(* IEC 61131-3 sources: plcassist-cli/packages/volt-lsp-iec/test-corpus/bakon-nano/Device/Plc Logic/Application/Library Manager/L_UBUP_BasicUtilities, 147 files *)

(* ---- L_UBUP_INTERNAL.gvl ---- *)
VAR_GLOBAL
	ONLINECHANGEDETECTION : L_UBUP_OnlineChangeDetection;
	LMJOBADMINSTRATION : L_UBUP_JobAdminstration;
	G_FBPOOLQUEUE : L_UBUP_JobPoolQueue;
	G_ILOWESTREQUESTPRIO : INT := DWORD_TO_INT(16#7FFF);
	G_DWCALLIDUNASSIGNED : DWORD := 4711;
	CDIENUMSTARTVALUE : DINT := 10000;
END_VAR

(* ---- L_UBUP_IACTIONPROVIDER.itf ---- *)
INTERFACE L_UBUP_IACTIONPROVIDER
END_INTERFACE

METHOD CYCLICACTION
VAR_INPUT
	ITFTIMINGCONTROLLER : L_UBUP_ITimingController;
END_VAR
VAR_OUTPUT
	XCOMPLETE : BOOL;
	XABORT : BOOL;
	IERRORID : INT;
END_VAR
END_METHOD

METHOD FINALIZEACTION
VAR_INPUT
	XABORTPROPOSED : BOOL;
	IERRORIDPROPOSED : INT;
END_VAR
VAR_OUTPUT
	XCOMPLETE : BOOL;
	XABORT : BOOL;
	IERRORID : INT;
END_VAR
END_METHOD

METHOD RESETACTION
VAR_OUTPUT
	XCOMPLETE : BOOL;
END_VAR
END_METHOD

METHOD STARTACTION
VAR_OUTPUT
	XCOMPLETE : BOOL;
	IERRORID : INT;
END_VAR
END_METHOD

(* ---- L_UBUP_IAFTERREADINPUTS.itf ---- *)
INTERFACE L_UBUP_IAFTERREADINPUTS
END_INTERFACE

METHOD AFTERREADINPUTS : INT
END_METHOD

(* ---- L_UBUP_IAFTERREADINPUTSEXIT.itf ---- *)
INTERFACE L_UBUP_IAFTERREADINPUTSEXIT
END_INTERFACE

METHOD AFTERREADINPUTSEXIT : INT
END_METHOD

(* ---- L_UBUP_IAFTERWRITEOUTPUTS.itf ---- *)
INTERFACE L_UBUP_IAFTERWRITEOUTPUTS
END_INTERFACE

METHOD AFTERWRITEOUTPUTS : INT
END_METHOD

(* ---- L_UBUP_IAFTERWRITEOUTPUTSEXIT.itf ---- *)
INTERFACE L_UBUP_IAFTERWRITEOUTPUTSEXIT
END_INTERFACE

METHOD AFTERWRITEOUTPUTSEXIT : INT
END_METHOD

(* ---- L_UBUP_IALLOCPOINTADRPROVIDER.itf ---- *)
INTERFACE L_UBUP_IALLOCPOINTADRPROVIDER
END_INTERFACE

METHOD ALLOCPOINTADR
VAR_OUTPUT
	IERRORID : INT;
END_VAR
END_METHOD

(* ---- L_UBUP_IALTERNATIVEREQUESTBYFAILEDCONDITION.itf ---- *)
INTERFACE L_UBUP_IALTERNATIVEREQUESTBYFAILEDCONDITION
END_INTERFACE

METHOD HANDLEREJECTEDREQUEST : BOOL
VAR_INPUT
	ITFREQUESTANNOUNCED : L_UBUP_IRequest;
END_VAR
VAR_OUTPUT
	ITFALTERNATIVEREQUEST : L_UBUP_IRequest;
END_VAR
END_METHOD

(* ---- L_UBUP_IBEFOREREADINPUTS.itf ---- *)
INTERFACE L_UBUP_IBEFOREREADINPUTS
END_INTERFACE

METHOD BEFOREREADINPUTS : INT
END_METHOD

(* ---- L_UBUP_IBEFOREREADINPUTSENTRY.itf ---- *)
INTERFACE L_UBUP_IBEFOREREADINPUTSENTRY
END_INTERFACE

METHOD BEFOREREADINPUTSENTRY : INT
END_METHOD

(* ---- L_UBUP_IBEFOREWRITEOUTPUTS.itf ---- *)
INTERFACE L_UBUP_IBEFOREWRITEOUTPUTS
END_INTERFACE

METHOD BEFOREWRITEOUTPUTS : INT
END_METHOD

(* ---- L_UBUP_IBEFOREWRITEOUTPUTSENTRY.itf ---- *)
INTERFACE L_UBUP_IBEFOREWRITEOUTPUTSENTRY
END_INTERFACE

METHOD BEFOREWRITEOUTPUTSENTRY : INT
END_METHOD

(* ---- L_UBUP_IBREAKPOINT.itf ---- *)
INTERFACE L_UBUP_IBREAKPOINT
END_INTERFACE

METHOD BREAKPOINT : INT
END_METHOD

(* ---- L_UBUP_ICATEGORY.itf ---- *)
INTERFACE L_UBUP_ICATEGORY
END_INTERFACE

METHOD CLASSIFY : BOOL
VAR_INPUT
	ECATEGORY : DINT;
END_VAR
END_METHOD

(* ---- L_UBUP_ICHECKER.itf ---- *)
INTERFACE L_UBUP_ICHECKER
END_INTERFACE

METHOD PERFORMCHECK : BOOL
VAR_INPUT
	WCONTEXT : DWORD;
END_VAR
END_METHOD

(* ---- L_UBUP_ICOMMAND.itf ---- *)
INTERFACE L_UBUP_ICOMMAND
END_INTERFACE

METHOD UPDATECOMMANDDATA : BOOL
VAR_INPUT
	DWCALLID : DWORD;
	XCONTINUOUSUPDATE : BOOL;
END_VAR
VAR_IN_OUT
	SCCOMMAND : L_UBUP_CommandData;
END_VAR
END_METHOD

(* ---- L_UBUP_ICOMPARER.itf ---- *)
INTERFACE L_UBUP_ICOMPARER
END_INTERFACE

METHOD COMPARE : DINT
VAR_INPUT
	DWARRIDX1 : DWORD;
	DWARRIDX2 : DWORD;
END_VAR
END_METHOD

(* ---- L_UBUP_ICONDITION.itf ---- *)
INTERFACE L_UBUP_ICONDITION
END_INTERFACE

METHOD VERIFY : BOOL
VAR_OUTPUT
	XCONDITIONERROR : BOOL;
	EERRORIDPROPOSED : L_IE1P_Error;
END_VAR
END_METHOD

(* ---- L_UBUP_ICRITICALSECTION.itf ---- *)
INTERFACE L_UBUP_ICRITICALSECTION
END_INTERFACE

METHOD LOCK : BOOL
END_METHOD

METHOD LOCKSTATE : BOOL
END_METHOD

METHOD UNLOCK : BOOL
END_METHOD

(* ---- L_UBUP_IEXCEPTION.itf ---- *)
INTERFACE L_UBUP_IEXCEPTION
END_INTERFACE

METHOD EXCEPTION : INT
END_METHOD

(* ---- L_UBUP_IFBPOOL.itf ---- *)
INTERFACE L_UBUP_IFBPOOL
END_INTERFACE

METHOD FREEINSTANCE : BOOL
VAR_INPUT
	ITFINSTANCE : L_UBUP_IPoolInstance;
	XWHANDLE : __XWORD;
END_VAR
END_METHOD

METHOD GETCAPACITY : BOOL
VAR_INPUT
	ECLASSID : DINT;
END_VAR
VAR_OUTPUT
	DWCAPACITY : DWORD;
END_VAR
END_METHOD

METHOD QUERYINSTANCE : BOOL
VAR_INPUT
	ECLASSID : DINT;
END_VAR
VAR_IN_OUT
	ITFINSTANCE : L_UBUP_IPoolInstance;
END_VAR
END_METHOD

(* ---- L_UBUP_IINSTANCE.itf ---- *)
INTERFACE L_UBUP_IINSTANCE
END_INTERFACE

(* ---- L_UBUP_IINSTANCELIST.itf ---- *)
INTERFACE L_UBUP_IINSTANCELIST
END_INTERFACE

METHOD APPENDPROXY : BOOL
VAR_INPUT
	ITFINSTANCELISTITEM : L_UBUP_IInstanceListProxy;
END_VAR
END_METHOD

(* ---- L_UBUP_IINSTANCELISTPASSENGER.itf ---- *)
INTERFACE L_UBUP_IINSTANCELISTPASSENGER
END_INTERFACE

(* ---- L_UBUP_IINSTANCELISTPROXY.itf ---- *)
INTERFACE L_UBUP_IINSTANCELISTPROXY
END_INTERFACE

(* ---- L_UBUP_IITERATOR.itf ---- *)
INTERFACE L_UBUP_IITERATOR
END_INTERFACE

METHOD NEXT : DWORD
END_METHOD

METHOD PREV : DWORD
END_METHOD

METHOD REWIND
VAR_OUTPUT
	DWARRAYIDXSTART : DWORD;
END_VAR
END_METHOD

(* ---- L_UBUP_IJOB.itf ---- *)
INTERFACE L_UBUP_IJOB
END_INTERFACE

METHOD EXPAND : BOOL
VAR_INPUT
	ITFSENDER : L_UBUP_ICommand;
	DWCALLID : DWORD;
END_VAR
VAR_OUTPUT
	EERRORID : L_IE1P_Error;
END_VAR
END_METHOD

METHOD HANDOVERRESOURCE : BOOL
VAR_INPUT
	ITFRESOURCE : L_UBUP_IUnknown;
END_VAR
END_METHOD

METHOD LINK : BOOL
VAR_INPUT
	ITFJOB : L_UBUP_IJob;
	XPREV : BOOL;
END_VAR
VAR_OUTPUT
	EERRORID : L_IE1P_Error;
END_VAR
END_METHOD

METHOD RELEASE
END_METHOD

(* ---- L_UBUP_IJOBACTION.itf ---- *)
INTERFACE L_UBUP_IJOBACTION
END_INTERFACE

METHOD ABORT
END_METHOD

METHOD CYCLE
VAR_OUTPUT
	ESTATE : L_UBUP_JobState;
	EERRORID : L_IE1P_Error;
END_VAR
END_METHOD

METHOD FINISH
END_METHOD

METHOD UPDATEREPORTDATA : BOOL
VAR_INPUT
	DWCALLID : DWORD;
END_VAR
VAR_IN_OUT
	SCREPORT : L_UBUP_ReportData;
END_VAR
END_METHOD

METHOD UPDATEREPORTRECEIVER : BOOL
VAR_INPUT
	ITFJOBREPORT : L_UBUP_IJobReport;
END_VAR
END_METHOD

(* ---- L_UBUP_IJOBCOLLECTION.itf ---- *)
INTERFACE L_UBUP_IJOBCOLLECTION
END_INTERFACE

METHOD GETJOB : BOOL
VAR_INPUT
	DWARRIDX : DWORD;
END_VAR
VAR_OUTPUT
	ITFJOB : L_UBUP_IJob;
END_VAR
END_METHOD

(* ---- L_UBUP_IJOBRECEIVER.itf ---- *)
INTERFACE L_UBUP_IJOBRECEIVER
END_INTERFACE

METHOD INSERT : BOOL
VAR_INPUT
	ITFJOB : L_UBUP_IJob;
END_VAR
END_METHOD

METHOD UNPLUGLISTENER : BOOL
VAR_INPUT
	ITFLISTENER : L_UBUP_IJobReceiverListener;
END_VAR
END_METHOD

METHOD ANNOUNCELISTENER : BOOL
VAR_INPUT
	ITFLISTENER : L_UBUP_IJobReceiverListener;
END_VAR
END_METHOD

(* ---- L_UBUP_IJOBRECEIVERLISTENER.itf ---- *)
INTERFACE L_UBUP_IJOBRECEIVERLISTENER
END_INTERFACE

METHOD LISTENAFTERCYCLE
VAR_INPUT
	ITFJOB : L_UBUP_IJob;
END_VAR
END_METHOD

METHOD LISTENINSERT
VAR_INPUT
	ITFJOB : L_UBUP_IJob;
	XSUCCEEDED : BOOL;
END_VAR
END_METHOD

(* ---- L_UBUP_IJOBREPORT.itf ---- *)
INTERFACE L_UBUP_IJOBREPORT
END_INTERFACE

METHOD RECEIVEREPORT
VAR_INPUT
	ITFJOB : L_UBUP_IJob;
END_VAR
END_METHOD

(* ---- L_UBUP_ILIST.itf ---- *)
INTERFACE L_UBUP_ILIST
END_INTERFACE

(* ---- L_UBUP_ILISTCONTROL.itf ---- *)
INTERFACE L_UBUP_ILISTCONTROL
END_INTERFACE

METHOD APPEND : BOOL
VAR_OUTPUT
	DWARRIDX : DWORD;
END_VAR
END_METHOD

METHOD GETARRIDXOF : DWORD
VAR_INPUT
	DWPOSITION : DWORD;
END_VAR
END_METHOD

METHOD GETMAX : DWORD
VAR_INPUT
	ITFCOMPARER : L_UBUP_IComparer;
END_VAR
END_METHOD

METHOD GETPOSITIONOF : DWORD
VAR_INPUT
	DWARRIDX : DWORD;
END_VAR
END_METHOD

METHOD INSERTAFTER : BOOL
VAR_INPUT
	DWARRIDX : DWORD;
END_VAR
VAR_OUTPUT
	DWNEXTIDX : DWORD;
END_VAR
END_METHOD

METHOD INSERTBEFORE : BOOL
VAR_INPUT
	DWARRIDX : DWORD;
END_VAR
VAR_OUTPUT
	DWPREVIDX : DWORD;
END_VAR
END_METHOD

METHOD REMOVE : BOOL
VAR_INPUT
	DWARRIDX : DWORD;
END_VAR
END_METHOD

METHOD SHIFTNEXT : BOOL
VAR_INPUT
	DWARRIDX : DWORD;
END_VAR
END_METHOD

METHOD SHIFTPREV : BOOL
VAR_INPUT
	DWARRIDX : DWORD;
END_VAR
END_METHOD

METHOD SORT : BOOL
VAR_INPUT
	ITFCOMPARER : L_UBUP_IComparer;
END_VAR
END_METHOD

METHOD SWAP : BOOL
VAR_INPUT
	DWARRIDX1 : DWORD;
	DWARRIDX2 : DWORD;
END_VAR
END_METHOD

METHOD TRYAPPEND : BOOL
VAR_INPUT
	DWARRIDX : DWORD;
END_VAR
END_METHOD

(* ---- L_UBUP_ILMDATA.itf ---- *)
INTERFACE L_UBUP_ILMDATA
END_INTERFACE

METHOD ABORT : UDINT
END_METHOD

METHOD EXECUTE : UDINT
END_METHOD

(* ---- L_UBUP_ILOCKABLE.itf ---- *)
INTERFACE L_UBUP_ILOCKABLE
END_INTERFACE

METHOD LOCK : BOOL
END_METHOD

METHOD LOCKSTATE : BOOL
END_METHOD

METHOD UNLOCK : BOOL
END_METHOD

(* ---- L_UBUP_IMAPOUTPUTSPROVIDER.itf ---- *)
INTERFACE L_UBUP_IMAPOUTPUTSPROVIDER
END_INTERFACE

METHOD MAPOUTPUTS
END_METHOD

(* ---- L_UBUP_IMAPSTATE.itf ---- *)
INTERFACE L_UBUP_IMAPSTATE
END_INTERFACE

(* ---- L_UBUP_IMEMORYCONSUMER.itf ---- *)
INTERFACE L_UBUP_IMEMORYCONSUMER
END_INTERFACE

METHOD EVALMEMORYPROVIDER
VAR_INPUT
	ITFMEMORYPROVIDER : L_UBUP_IMemoryProvider;
END_VAR
END_METHOD

(* ---- L_UBUP_IMEMORYPROVIDER.itf ---- *)
INTERFACE L_UBUP_IMEMORYPROVIDER
END_INTERFACE

METHOD REGISTERCONSUMER
VAR_INPUT
	ITFMEMORYCONSUMER : L_UBUP_IMemoryConsumer;
END_VAR
END_METHOD

(* ---- L_UBUP_IMONITORSTATESERVER.itf ---- *)
INTERFACE L_UBUP_IMONITORSTATESERVER
END_INTERFACE

METHOD MONITORCASE
VAR_INPUT
	ECASE : L_UBUP_StateHandleCase;
END_VAR
END_METHOD

METHOD MONITORREQUEST : INT
VAR_INPUT
	ITFREQUEST : L_UBUP_IRequest;
END_VAR
END_METHOD

METHOD MONITORREQUESTANNOUNCED : INT
VAR_INPUT
	ITFREQUESTANNOUNCED : L_UBUP_IRequest;
	ITFREQUESTALTERNATIVE : L_UBUP_IRequest := 0;
	ITFREQUESTACTIVE : L_UBUP_IRequest;
END_VAR
END_METHOD

(* ---- L_UBUP_IOBJECT.itf ---- *)
INTERFACE L_UBUP_IOBJECT
END_INTERFACE

METHOD CALL_INIT : BOOL
END_METHOD

METHOD SETNEXT : BOOL
VAR_INPUT
	ITFOBJECT : L_UBUP_IObject;
END_VAR
END_METHOD

METHOD SETPREV : BOOL
VAR_INPUT
	ITFOBJECT : L_UBUP_IObject;
END_VAR
END_METHOD

(* ---- L_UBUP_IOBJECTQUEUE.itf ---- *)
INTERFACE L_UBUP_IOBJECTQUEUE
END_INTERFACE

METHOD DEQUEUE : BOOL
END_METHOD

METHOD ENQUEUE : BOOL
VAR_INPUT
	ITFOBJECT : L_UBUP_IObject;
END_VAR
END_METHOD

METHOD REMOVE : BOOL
VAR_INPUT
	ITFOBJECT : L_UBUP_IObject;
END_VAR
END_METHOD

(* ---- L_UBUP_IPLCOPENSTATUS.itf ---- *)
INTERFACE L_UBUP_IPLCOPENSTATUS
END_INTERFACE

METHOD GET_EERRORID : L_IE1P_Error
END_METHOD

METHOD GET_XACTIVE : BOOL
END_METHOD

METHOD GET_XBUSY : BOOL
END_METHOD

METHOD GET_XCOMMANDABORTED : BOOL
END_METHOD

METHOD GET_XDONE : BOOL
END_METHOD

METHOD GET_XINITIAL : BOOL
END_METHOD

(* ---- L_UBUP_IPOINTERCOLLECTION.itf ---- *)
INTERFACE L_UBUP_IPOINTERCOLLECTION
END_INTERFACE

METHOD GETPOINTER : BOOL
VAR_INPUT
	DWARRIDX : DWORD;
END_VAR
VAR_OUTPUT
	PBYTE : POINTER TO BYTE;
END_VAR
END_METHOD

(* ---- L_UBUP_IPOOLINSTANCE.itf ---- *)
INTERFACE L_UBUP_IPOOLINSTANCE
END_INTERFACE

METHOD FREE : BOOL
END_METHOD

METHOD OCCUPY : BOOL
VAR_INPUT
	ITFOWNER : L_UBUP_IFBPool;
	XWHANDLE : __XWORD;
END_VAR
END_METHOD

(* ---- L_UBUP_IQUEUE.itf ---- *)
INTERFACE L_UBUP_IQUEUE
END_INTERFACE

METHOD DEQUEUE : BOOL
END_METHOD

METHOD ENQUEUE : BOOL
END_METHOD

METHOD GETEMPTY : BOOL
VAR_OUTPUT
	PBYTE : POINTER TO BYTE;
	DWSIZE : DWORD;
END_VAR
END_METHOD

METHOD GETPEEK : BOOL
VAR_OUTPUT
	PBYTE : POINTER TO BYTE;
	DWSIZE : DWORD;
END_VAR
END_METHOD

METHOD RESET : BOOL
END_METHOD

(* ---- L_UBUP_IREADINPUTSEXIT.itf ---- *)
INTERFACE L_UBUP_IREADINPUTSEXIT
END_INTERFACE

METHOD READINPUTSEXIT : INT
END_METHOD

(* ---- L_UBUP_IREFCOUNTER.itf ---- *)
INTERFACE L_UBUP_IREFCOUNTER
END_INTERFACE

METHOD DECCOUNTER : DINT
END_METHOD

METHOD INCCOUNTER : DINT
END_METHOD

(* ---- L_UBUP_IREQUEST.itf ---- *)
INTERFACE L_UBUP_IREQUEST
END_INTERFACE

METHOD CONFIRM : INT
VAR_IN_OUT
	IREQUEST : L_UBUP_IRequest;
END_VAR
END_METHOD

METHOD FORCESTATEENTRY : BOOL
END_METHOD

(* ---- L_UBUP_ISTATECLIENT.itf ---- *)
INTERFACE L_UBUP_ISTATECLIENT
END_INTERFACE

METHOD CALLFBS
VAR_INPUT
	ECASE : L_UBUP_StateHandleCase;
END_VAR
END_METHOD

METHOD CALLSTATE
VAR_INPUT
	ITFSTATESERVER : L_UBUP_IStateServer;
	ISTATE : INT;
	ECASE : L_UBUP_StateHandleCase;
END_VAR
END_METHOD

METHOD CHECKTRANSITION
VAR_INPUT
	ITFSTATESERVER : L_UBUP_IStateServer;
END_VAR
END_METHOD

METHOD DISABLECLIENT : BOOL
VAR_INPUT
	XFIRSTCALL : BOOL;
END_VAR
END_METHOD

METHOD ENABLECLIENT : BOOL
VAR_INPUT
	XFIRSTCALL : BOOL;
END_VAR
END_METHOD

METHOD FINALIZECYCLE
END_METHOD

METHOD LEAVESTATE
END_METHOD

METHOD PREPARECYCLE
END_METHOD

METHOD PREPARESTATECHANGE
END_METHOD

METHOD STIMULATETRANSITION
VAR_INPUT
	ECASE : L_UBUP_StateHandleCase;
END_VAR
END_METHOD

METHOD UPDATECONDITIONERROR : BOOL
VAR_INPUT
	ITFREQUEST : L_UBUP_IRequest;
END_VAR
END_METHOD

(* ---- L_UBUP_ISTATECLIENTDECORATOR.itf ---- *)
INTERFACE L_UBUP_ISTATECLIENTDECORATOR
END_INTERFACE

METHOD EXTENDEDCALLFBS
VAR_INPUT
	ECASE : L_UBUP_StateHandleCase;
END_VAR
END_METHOD

METHOD EXTENDEDCALLSTATE
VAR_INPUT
	ITFBASE : L_UBUP_IStateClient;
	ITFSTATESERVER : L_UBUP_IStateServer;
	ISTATE : INT;
	ECASE : L_UBUP_StateHandleCase;
END_VAR
END_METHOD

METHOD EXTENDEDCHECKTRANSITION
VAR_INPUT
	ITFSTATESERVER : L_UBUP_IStateServer;
END_VAR
END_METHOD

METHOD EXTENDEDDISABLECLIENT : BOOL
VAR_INPUT
	XFIRSTCALL : BOOL;
END_VAR
END_METHOD

METHOD EXTENDEDENABLECLIENT : BOOL
VAR_INPUT
	XFIRSTCALL : BOOL;
END_VAR
END_METHOD

METHOD EXTENDEDFINALIZECYCLE
END_METHOD

METHOD EXTENDEDPREPARECYCLE
END_METHOD

METHOD EXTENDEDPREPARESTATECHANGE
END_METHOD

METHOD EXTENDEDSTIMULATETRANSITION
VAR_INPUT
	ECASE : L_UBUP_StateHandleCase;
END_VAR
END_METHOD

(* ---- L_UBUP_ISTATESERVER.itf ---- *)
INTERFACE L_UBUP_ISTATESERVER
END_INTERFACE

METHOD ANNOUNCENEWREQUEST
END_METHOD

METHOD FREEZEREQUEST
VAR_INPUT
	EERRORIDBYBLOCKEFREEZEREQUEST : L_IE1P_Error;
END_VAR
END_METHOD

METHOD ISACTIVE : BOOL
VAR_INPUT
	ITFREQUEST : L_UBUP_IRequest;
END_VAR
END_METHOD

METHOD REQUESTS : INT
VAR_INPUT
	ITFREQUEST : L_UBUP_IRequest;
END_VAR
END_METHOD

METHOD UNFREEZEREQUEST : BOOL
END_METHOD

METHOD VERIFYFREEZEREQUEST : BOOL
VAR_INPUT
	ITFREQUEST : L_UBUP_IRequest;
END_VAR
VAR_OUTPUT
	XCONDITIONERROR : BOOL;
	EERRORIDPROPOSED : L_IE1P_Error;
END_VAR
END_METHOD

(* ---- L_UBUP_ISTRINGCOLLECTION.itf ---- *)
INTERFACE L_UBUP_ISTRINGCOLLECTION
END_INTERFACE

METHOD GETSTRING : BOOL
VAR_INPUT
	DWARRIDX : DWORD;
END_VAR
VAR_OUTPUT
	STVALUE : STRING(255);
END_VAR
END_METHOD

(* ---- L_UBUP_ITIMINGCONTROLLER.itf ---- *)
INTERFACE L_UBUP_ITIMINGCONTROLLER
END_INTERFACE

METHOD CHECKTIMING
VAR_OUTPUT
	XTIMEOUT : BOOL;
	XTIMELIMIT : BOOL;
END_VAR
END_METHOD

METHOD STARTINVOCATIONTIMER
END_METHOD

METHOD STARTOPERATIONTIMER
END_METHOD

(* ---- L_UBUP_IUNKNOWN.itf ---- *)
INTERFACE L_UBUP_IUNKNOWN
END_INTERFACE

METHOD REQUESTINTERFACE : BOOL
VAR_INPUT
	ID : DINT;
	PITFUNKNOWN : POINTER TO L_UBUP_IUnknown;
END_VAR
END_METHOD

(* ---- L_UBUP_IWRITEOUTPUTSENTRY.itf ---- *)
INTERFACE L_UBUP_IWRITEOUTPUTSENTRY
END_INTERFACE

METHOD WRITEOUTPUTSENTRY : INT
END_METHOD

(* ---- GETBOOLEANPROPERTY.fun ---- *)
FUNCTION GETBOOLEANPROPERTY : BOOL
VAR_INPUT
	STKEY : WSTRING;
END_VAR
END_FUNCTION

(* ---- GETCOMPANY.fun ---- *)
FUNCTION GETCOMPANY : WSTRING
END_FUNCTION

(* ---- GETNUMBERPROPERTY.fun ---- *)
FUNCTION GETNUMBERPROPERTY : DINT
VAR_INPUT
	STKEY : WSTRING;
END_VAR
END_FUNCTION

(* ---- GETTEXTPROPERTY.fun ---- *)
FUNCTION GETTEXTPROPERTY : WSTRING
VAR_INPUT
	STKEY : WSTRING;
END_VAR
END_FUNCTION

(* ---- GETTEXTPROPERTY2.fun ---- *)
FUNCTION GETTEXTPROPERTY2 : POINTER TO WSTRING
VAR_INPUT
	STKEY : WSTRING;
END_VAR
END_FUNCTION

(* ---- GETTITLE.fun ---- *)
FUNCTION GETTITLE : WSTRING
END_FUNCTION

(* ---- GETVERSION.fun ---- *)
FUNCTION GETVERSION : VERSION
END_FUNCTION

(* ---- GETVERSIONPROPERTY.fun ---- *)
FUNCTION GETVERSIONPROPERTY : VERSION
VAR_INPUT
	STKEY : WSTRING;
END_VAR
END_FUNCTION

(* ---- L_UBUP_CREATECALLID.fun ---- *)
FUNCTION L_UBUP_CREATECALLID : DWORD
END_FUNCTION

(* ---- L_UBUP_CREATEOBJECTID.fun ---- *)
FUNCTION L_UBUP_CREATEOBJECTID : DWORD
END_FUNCTION

(* ---- L_UBUP_FILEADDRESS.fun ---- *)
FUNCTION L_UBUP_FILEADDRESS : STRING(255)
END_FUNCTION

(* ---- L_UBUP_GETTASKCYCLE.fun ---- *)
FUNCTION L_UBUP_GETTASKCYCLE : LREAL
VAR_INPUT
	LRCYCLETIMEIN : LREAL;
END_VAR
END_FUNCTION

(* ---- L_UBUP_GETTASKINFO.fun ---- *)
FUNCTION L_UBUP_GETTASKINFO : BOOL
VAR_OUTPUT
	ITASKINDEX : INT;
	HTASK : RTS_IEC_HANDLE;
	HIECTASK : RTS_IEC_HANDLE;
	PSCSYSTASKINFO : POINTER TO SYS_TASK_INFO;
	UDIOSPRIORITY : UDINT;
	UDIPRIORITY : UDINT;
	UDITASKINTERVAL : UDINT;
END_VAR
END_FUNCTION

(* ---- L_UBUP_ISLENZETARGET.fun ---- *)
FUNCTION L_UBUP_ISLENZETARGET : BOOL
VAR_OUTPUT
	DWVENDORID : DWORD;
END_VAR
END_FUNCTION

(* ---- L_UBUP_ISONLINECHANGEACTIVE.fun ---- *)
FUNCTION L_UBUP_ISONLINECHANGEACTIVE : BOOL
END_FUNCTION

(* ---- L_UBUP_LMDATAMANAGERINSERTDATA.fun ---- *)
FUNCTION L_UBUP_LMDATAMANAGERINSERTDATA : BOOL
VAR_INPUT
	ITFLMDATA : L_UBUP_ILMData;
END_VAR
END_FUNCTION

(* ---- L_UBUP_LOCALDATEANDTIME.fun ---- *)
FUNCTION L_UBUP_LOCALDATEANDTIME : BOOL
VAR_OUTPUT
	UIYEAR : UINT;
	UIMONTH : UINT;
	UIDAY : UINT;
	UIHOUR : UINT;
	UIMINUTE : UINT;
	UISECOND : UINT;
	UIMILLISECONDS : UINT;
	UIWEEKDAY : UINT;
	DATDATE : DATE;
	TODTIME : TIME_OF_DAY;
END_VAR
END_FUNCTION

(* ---- L_UBUP_QUERY_IJOB_ALL.fun ---- *)
FUNCTION L_UBUP_QUERY_IJOB_ALL : BOOL
VAR_INPUT
	ITFJOB : L_UBUP_IJob;
END_VAR
VAR_OUTPUT
	ITFINSTANCE : L_UBUP_IPoolInstance;
	ITFSTATECLIENT : L_UBUP_IStateClient;
	ITFPLCOPENSTATUS : L_UBUP_IPLCOpenStatus;
END_VAR
END_FUNCTION

(* ---- L_UBUP_QUERY_IJOB_IINSTANCE.fun ---- *)
FUNCTION L_UBUP_QUERY_IJOB_IINSTANCE : BOOL
VAR_INPUT
	ITFJOB : L_UBUP_IJob;
END_VAR
VAR_OUTPUT
	ITFINSTANCE : L_UBUP_IPoolInstance;
END_VAR
END_FUNCTION

(* ---- L_UBUP_QUERY_IJOB_IPLCOPENSTATUS.fun ---- *)
FUNCTION L_UBUP_QUERY_IJOB_IPLCOPENSTATUS : BOOL
VAR_INPUT
	ITFJOB : L_UBUP_IJob;
END_VAR
VAR_OUTPUT
	ITFPLCOPENSTATUS : L_UBUP_IPLCOpenStatus;
END_VAR
END_FUNCTION

(* ---- L_UBUP_SYMBOLCONFIGREADNUMVAR.fun ---- *)
FUNCTION L_UBUP_SYMBOLCONFIGREADNUMVAR : BOOL
VAR_INPUT
	SVARIABLENAME : STRING;
END_VAR
VAR_OUTPUT
	SCVARIABLE : L_UBUP_Variable;
END_VAR
END_FUNCTION

(* ---- L_UBUP_SYMBOLCONFIGREADSTRINGVAR.fun ---- *)
FUNCTION L_UBUP_SYMBOLCONFIGREADSTRINGVAR : BOOL
VAR_INPUT
	SVARIABLENAME : STRING;
END_VAR
VAR_OUTPUT
	SVALUE : STRING;
END_VAR
END_FUNCTION

(* ---- L_UBUP_SYMBOLCONFIGREADVAR.fun ---- *)
FUNCTION L_UBUP_SYMBOLCONFIGREADVAR : BOOL
VAR_INPUT
	SVARIABLENAME : STRING;
END_VAR
VAR_OUTPUT
	SCVARIABLE : L_UBUP_Variable;
END_VAR
END_FUNCTION

(* ---- L_UBUP_SYMBOLCONFIGREADVARASDWORD.fun ---- *)
FUNCTION L_UBUP_SYMBOLCONFIGREADVARASDWORD : BOOL
VAR_INPUT
	SVARIABLENAME : STRING;
END_VAR
VAR_OUTPUT
	DWVALUE : DWORD;
END_VAR
END_FUNCTION

(* ---- L_UBUP_SYMBOLCONFIGREADVARASLINT.fun ---- *)
FUNCTION L_UBUP_SYMBOLCONFIGREADVARASLINT : BOOL
VAR_INPUT
	SVARIABLENAME : STRING;
END_VAR
VAR_OUTPUT
	LIVALUE : LINT;
END_VAR
END_FUNCTION

(* ---- L_UBUP_SYMBOLCONFIGREADVARASLREAL.fun ---- *)
FUNCTION L_UBUP_SYMBOLCONFIGREADVARASLREAL : BOOL
VAR_INPUT
	SVARIABLENAME : STRING;
END_VAR
VAR_OUTPUT
	LRVALUE : LREAL;
END_VAR
END_FUNCTION

(* ---- L_UBUP_SYMBOLCONFIGREADVARASWORD.fun ---- *)
FUNCTION L_UBUP_SYMBOLCONFIGREADVARASWORD : BOOL
VAR_INPUT
	SVARIABLENAME : STRING;
END_VAR
VAR_OUTPUT
	WVALUE : WORD;
END_VAR
END_FUNCTION

(* ---- L_UBUP_SYMBOLCONFIGSYMBOLEXISTS.fun ---- *)
FUNCTION L_UBUP_SYMBOLCONFIGSYMBOLEXISTS : BOOL
VAR_INPUT
	SVARIABLENAME : STRING;
END_VAR
END_FUNCTION

(* ---- GLOBALTEXTLIST.fb ---- *)
FUNCTION_BLOCK GLOBALTEXTLIST
VAR
	M_TEXTLISTFILE : STRING(255);
	_STNAMESPACE : STRING;
END_VAR
END_FUNCTION_BLOCK

(* ---- L_UBUP_BEHAVIOURMODEL.fb ---- *)
FUNCTION_BLOCK L_UBUP_BEHAVIOURMODEL
VAR_INPUT
	XCONTROL : BOOL;
	XABORT : BOOL;
	UDITIMELIMIT : SYSTIME;
	UDITIMEOUT : SYSTIME;
END_VAR
VAR_OUTPUT
	XDONE : BOOL;
	XBUSY : BOOL;
	XABORTED : BOOL;
	XERROR : BOOL;
	IERRORID : INT;
END_VAR
VAR
	ITFAP : L_UBUP_IActionProvider;
	ITFTC : L_UBUP_ITimingController;
	ITFADR : L_UBUP_IAllocPointAdrProvider;
	ITFMAP : L_UBUP_IMapOutputsProvider;
	_ESTATE : L_UBUP_BehaviourModelState := L_UBUP_BehaviourModelState.DORMANT;
	_IERRORIDPROPOSED : INT;
	_XRESETREQUEST : BOOL;
	BEHAVIOURMODELTYPE : L_UBUP_BehaviourModelType;
END_VAR
END_FUNCTION_BLOCK

METHOD HANDLEABORTEDSTATE
VAR_OUTPUT
	XAGAIN : BOOL;
END_VAR
VAR_IN_OUT
	ESTATE : L_UBUP_BehaviourModelState;
END_VAR
END_METHOD

METHOD HANDLEABORTINGSTATE
VAR_OUTPUT
	XAGAIN : BOOL;
END_VAR
VAR_IN_OUT
	ESTATE : L_UBUP_BehaviourModelState;
END_VAR
END_METHOD

METHOD HANDLECLEANINGSTATE
VAR_OUTPUT
	XAGAIN : BOOL;
END_VAR
VAR_IN_OUT
	ESTATE : L_UBUP_BehaviourModelState;
END_VAR
END_METHOD

METHOD HANDLEDONESTATE
VAR_OUTPUT
	XAGAIN : BOOL;
END_VAR
VAR_IN_OUT
	ESTATE : L_UBUP_BehaviourModelState;
END_VAR
END_METHOD

METHOD HANDLEDORMANTSTATE
VAR_OUTPUT
	XAGAIN : BOOL;
END_VAR
VAR_IN_OUT
	ESTATE : L_UBUP_BehaviourModelState;
END_VAR
END_METHOD

METHOD HANDLEERRORSTATE
VAR_OUTPUT
	XAGAIN : BOOL;
END_VAR
VAR_IN_OUT
	ESTATE : L_UBUP_BehaviourModelState;
END_VAR
END_METHOD

METHOD HANDLEEXECUTINGSTATE
VAR_OUTPUT
	XAGAIN : BOOL;
END_VAR
VAR_IN_OUT
	ESTATE : L_UBUP_BehaviourModelState;
END_VAR
END_METHOD

METHOD HANDLERESETTINGSTATE
VAR_OUTPUT
	XAGAIN : BOOL;
END_VAR
VAR_IN_OUT
	ESTATE : L_UBUP_BehaviourModelState;
END_VAR
END_METHOD

METHOD HANDLESTARTINGSTATE
VAR_OUTPUT
	XAGAIN : BOOL;
END_VAR
VAR_IN_OUT
	ESTATE : L_UBUP_BehaviourModelState;
END_VAR
END_METHOD

METHOD STATEMACHINE
VAR_IN_OUT
	ESTATE : L_UBUP_BehaviourModelState;
END_VAR
END_METHOD

METHOD FB_INIT : BOOL
VAR_INPUT
	BINITRETAINS : BOOL;
	BINCOPYCODE : BOOL;
	ITFAP : L_UBUP_IActionProvider;
END_VAR
END_METHOD

(* ---- L_UBUP_BEHAVIOURMODEL_ETRIG.fb ---- *)
FUNCTION_BLOCK L_UBUP_BEHAVIOURMODEL_ETRIG EXTENDS L_UBUP_BehaviourModel
VAR
	BEHAVIOURMODELTYPE : L_UBUP_BehaviourModelType;
END_VAR
END_FUNCTION_BLOCK

METHOD HANDLEEXECUTINGSTATE
VAR_OUTPUT
	XAGAIN : BOOL;
END_VAR
VAR_IN_OUT
	ESTATE : L_UBUP_BehaviourModelState;
END_VAR
END_METHOD

(* ---- L_UBUP_BEHAVIOURMODEL_ETRIGA.fb ---- *)
FUNCTION_BLOCK L_UBUP_BEHAVIOURMODEL_ETRIGA EXTENDS L_UBUP_BehaviourModel
VAR
	BEHAVIOURMODELTYPE : L_UBUP_BehaviourModelType;
END_VAR
END_FUNCTION_BLOCK

METHOD HANDLEEXECUTINGSTATE
VAR_OUTPUT
	XAGAIN : BOOL;
END_VAR
VAR_IN_OUT
	ESTATE : L_UBUP_BehaviourModelState;
END_VAR
END_METHOD

METHOD HANDLESTARTINGSTATE
VAR_OUTPUT
	XAGAIN : BOOL;
END_VAR
VAR_IN_OUT
	ESTATE : L_UBUP_BehaviourModelState;
END_VAR
END_METHOD

(* ---- L_UBUP_BEHAVIOURMODEL_ETRIGTO.fb ---- *)
FUNCTION_BLOCK L_UBUP_BEHAVIOURMODEL_ETRIGTO EXTENDS L_UBUP_BehaviourModelTC
VAR
	BEHAVIOURMODELTYPE : L_UBUP_BehaviourModelType;
END_VAR
END_FUNCTION_BLOCK

METHOD HANDLEEXECUTINGSTATE
VAR_OUTPUT
	XAGAIN : BOOL;
END_VAR
VAR_IN_OUT
	ESTATE : L_UBUP_BehaviourModelState;
END_VAR
END_METHOD

METHOD HANDLESTARTINGSTATE
VAR_OUTPUT
	XAGAIN : BOOL;
END_VAR
VAR_IN_OUT
	ESTATE : L_UBUP_BehaviourModelState;
END_VAR
END_METHOD

(* ---- L_UBUP_BEHAVIOURMODEL_LCON.fb ---- *)
FUNCTION_BLOCK L_UBUP_BEHAVIOURMODEL_LCON EXTENDS L_UBUP_BehaviourModel
VAR
	BEHAVIOURMODELTYPE : L_UBUP_BehaviourModelType;
END_VAR
END_FUNCTION_BLOCK

METHOD HANDLEEXECUTINGSTATE
VAR_OUTPUT
	XAGAIN : BOOL;
END_VAR
VAR_IN_OUT
	ESTATE : L_UBUP_BehaviourModelState;
END_VAR
END_METHOD

(* ---- L_UBUP_BEHAVIOURMODEL_LCONC.fb ---- *)
FUNCTION_BLOCK L_UBUP_BEHAVIOURMODEL_LCONC EXTENDS L_UBUP_BehaviourModel
VAR
	BEHAVIOURMODELTYPE : L_UBUP_BehaviourModelType;
END_VAR
END_FUNCTION_BLOCK

METHOD HANDLEDONESTATE
VAR_OUTPUT
	XAGAIN : BOOL;
END_VAR
VAR_IN_OUT
	ESTATE : L_UBUP_BehaviourModelState;
END_VAR
END_METHOD

METHOD HANDLEEXECUTINGSTATE
VAR_OUTPUT
	XAGAIN : BOOL;
END_VAR
VAR_IN_OUT
	ESTATE : L_UBUP_BehaviourModelState;
END_VAR
END_METHOD

(* ---- L_UBUP_BEHAVIOURMODEL_LCONC_LENZE.fb ---- *)
FUNCTION_BLOCK L_UBUP_BEHAVIOURMODEL_LCONC_LENZE EXTENDS L_UBUP_BehaviourModel
VAR
	BEHAVIOURMODELTYPE : L_UBUP_BehaviourModelType;
END_VAR
END_FUNCTION_BLOCK

METHOD HANDLEDONESTATE
VAR_OUTPUT
	XAGAIN : BOOL;
END_VAR
VAR_IN_OUT
	ESTATE : L_UBUP_BehaviourModelState;
END_VAR
END_METHOD

METHOD HANDLEEXECUTINGSTATE
VAR_OUTPUT
	XAGAIN : BOOL;
END_VAR
VAR_IN_OUT
	ESTATE : L_UBUP_BehaviourModelState;
END_VAR
END_METHOD

(* ---- L_UBUP_BEHAVIOURMODEL_LCONTO.fb ---- *)
FUNCTION_BLOCK L_UBUP_BEHAVIOURMODEL_LCONTO EXTENDS L_UBUP_BehaviourModelTC
VAR
	BEHAVIOURMODELTYPE : L_UBUP_BehaviourModelType;
END_VAR
END_FUNCTION_BLOCK

METHOD HANDLEEXECUTINGSTATE
VAR_OUTPUT
	XAGAIN : BOOL;
END_VAR
VAR_IN_OUT
	ESTATE : L_UBUP_BehaviourModelState;
END_VAR
END_METHOD

METHOD HANDLESTARTINGSTATE
VAR_OUTPUT
	XAGAIN : BOOL;
END_VAR
VAR_IN_OUT
	ESTATE : L_UBUP_BehaviourModelState;
END_VAR
END_METHOD

(* ---- L_UBUP_BEHAVIOURMODELTC.fb ---- *)
FUNCTION_BLOCK L_UBUP_BEHAVIOURMODELTC EXTENDS L_UBUP_BehaviourModel
END_FUNCTION_BLOCK

METHOD HANDLEDORMANTSTATE
VAR_OUTPUT
	XAGAIN : BOOL;
END_VAR
VAR_IN_OUT
	ESTATE : L_UBUP_BehaviourModelState;
END_VAR
END_METHOD

METHOD FB_INIT : BOOL
VAR_INPUT
	BINITRETAINS : BOOL;
	BINCOPYCODE : BOOL;
	ITFAP : L_UBUP_IActionProvider;
	ITFTC : L_UBUP_ITimingController;
END_VAR
END_METHOD

(* ---- L_UBUP_COMMANDSENDER.fb ---- *)
FUNCTION_BLOCK L_UBUP_COMMANDSENDER
VAR_INPUT
	XEXECUTE : BOOL;
	XREPORT : BOOL := TRUE;
	ITFREPORT : L_UBUP_IJobReport;
END_VAR
VAR_OUTPUT
	XCMDACCEPTED : BOOL;
	XDONE : BOOL;
	XBUSY : BOOL;
	XACTIVE : BOOL;
	XCOMMANDABORTED : BOOL;
	XERROR : BOOL;
	EERRORID : L_IE1P_Error;
	DWCALLID : DWORD := L_UBUP_Internal.g_dwCallIDUnassigned;
	ITFJOB : L_UBUP_IJob;
END_VAR
VAR
	_ECOMMANDTYPE : L_UBUP_CommandType;
	_PREPORT : POINTER TO L_UBUP_ReportData;
	_XREPORTVALID : BOOL;
	_XCYCLICSLAVE : BOOL;
	_ITFJOBPOOL : L_UBUP_IFBPool;
	_ITFJOBRECEIVER : L_UBUP_IJobReceiver;
	_ITFACTUALJOB : L_UBUP_IJob;
	_MODEL : L_UBUP_BehaviourModel_ETrigA;
	JOBCLASSID : DINT;
END_VAR
END_FUNCTION_BLOCK

METHOD CYCLICACTION
VAR_INPUT
	ITFTIMINGCONTROLLER : L_UBUP_ITimingController;
END_VAR
VAR_OUTPUT
	XCOMPLETE : BOOL;
	XABORT : BOOL;
	IERRORID : INT;
END_VAR
END_METHOD

METHOD FINALIZEACTION
VAR_INPUT
	XABORTPROPOSED : BOOL;
	IERRORIDPROPOSED : INT;
END_VAR
VAR_OUTPUT
	XCOMPLETE : BOOL;
	XABORT : BOOL;
	IERRORID : INT;
END_VAR
END_METHOD

METHOD RESETACTION
VAR_OUTPUT
	XCOMPLETE : BOOL;
END_VAR
END_METHOD

METHOD STARTACTION
VAR_OUTPUT
	XCOMPLETE : BOOL;
	IERRORID : INT;
END_VAR
END_METHOD

METHOD ALLOCPOINTADR
VAR_OUTPUT
	IERRORID : INT;
END_VAR
END_METHOD

METHOD UPDATECOMMANDDATA : BOOL
VAR_INPUT
	DWCALLID : DWORD;
	XCONTINUOUSUPDATE : BOOL;
END_VAR
VAR_IN_OUT
	SCCOMMAND : L_UBUP_CommandData;
END_VAR
END_METHOD

METHOD RECEIVEREPORT
VAR_INPUT
	ITFJOB : L_UBUP_IJob;
END_VAR
END_METHOD

METHOD REQUESTINTERFACE : BOOL
VAR_INPUT
	ID : DINT;
	PITFUNKNOWN : POINTER TO L_UBUP_IUnknown;
END_VAR
END_METHOD

METHOD FB_INIT : BOOL
VAR_INPUT
	BINITRETAINS : BOOL;
	BINCOPYCODE : BOOL;
END_VAR
END_METHOD

METHOD CALLERRORHANDLER
VAR_INPUT
	EERRORID : L_IE1P_Error;
END_VAR
END_METHOD

METHOD CHECKCMDACCEPTED : BOOL
END_METHOD

METHOD CONNECTJOB : BOOL
VAR_INPUT
	ITFJOBPOOL : L_UBUP_IFBPool;
END_VAR
VAR_OUTPUT
	ITFJOB : L_UBUP_IJob;
END_VAR
END_METHOD

METHOD CONNECTJOBPOOL : BOOL
END_METHOD

METHOD CONNECTJOBRECEIVER
END_METHOD

METHOD PREPARECYCLE
END_METHOD

METHOD REPORT2OUTPUTS
VAR_INPUT
	XRESET : BOOL;
END_VAR
END_METHOD

(* ---- L_UBUP_CONDITIONBASE.fb ---- *)
FUNCTION_BLOCK L_UBUP_CONDITIONBASE
VAR_OUTPUT
	XVERIFY : BOOL;
END_VAR
VAR
	XCALLVERIFY : BOOL;
	XCONDITIONERROR : BOOL;
	EERRORIDPROPOSED : L_IE1P_Error;
END_VAR
END_FUNCTION_BLOCK

METHOD VERIFY : BOOL
VAR_OUTPUT
	XCONDITIONERROR : BOOL;
	EERRORIDPROPOSED : L_IE1P_Error;
END_VAR
END_METHOD

(* ---- L_UBUP_CONDITIONCOLLECTION.fb ---- *)
FUNCTION_BLOCK L_UBUP_CONDITIONCOLLECTION EXTENDS L_UBUP_ConditionCollectionAND
END_FUNCTION_BLOCK

(* ---- L_UBUP_CONDITIONCOLLECTIONAND.fb ---- *)
FUNCTION_BLOCK L_UBUP_CONDITIONCOLLECTIONAND
VAR_INPUT
	AITFCONDITION : ARRAY [1..100] OF L_UBUP_ICondition;
END_VAR
VAR
	_IDX : INT;
END_VAR
END_FUNCTION_BLOCK

METHOD VERIFY : BOOL
VAR_OUTPUT
	XCONDITIONERROR : BOOL;
	EERRORIDPROPOSED : L_IE1P_Error;
END_VAR
END_METHOD

(* ---- L_UBUP_CONDITIONCOLLECTIONOR.fb ---- *)
FUNCTION_BLOCK L_UBUP_CONDITIONCOLLECTIONOR
VAR_INPUT
	AITFCONDITION : ARRAY [1..100] OF L_UBUP_ICondition;
END_VAR
VAR
	_IDX : INT;
END_VAR
END_FUNCTION_BLOCK

METHOD VERIFY : BOOL
VAR_OUTPUT
	XCONDITIONERROR : BOOL;
	EERRORIDPROPOSED : L_IE1P_Error;
END_VAR
END_METHOD

(* ---- L_UBUP_CONDITIONINPUT.fb ---- *)
FUNCTION_BLOCK L_UBUP_CONDITIONINPUT EXTENDS L_UBUP_ConditionBase
VAR_INPUT
	XCONDITION : BOOL;
END_VAR
VAR
	ECONDITIONWARNINGID_INT : L_IE1P_Error;
END_VAR
END_FUNCTION_BLOCK

METHOD VERIFY : BOOL
VAR_OUTPUT
	XCONDITIONERROR : BOOL;
	EERRORIDPROPOSED : L_IE1P_Error;
END_VAR
END_METHOD

METHOD FB_INIT : BOOL
VAR_INPUT
	BINITRETAINS : BOOL;
	BINCOPYCODE : BOOL;
	ECONDITIONWARNINGID : L_IE1P_Error;
END_VAR
END_METHOD

(* ---- L_UBUP_CONDITIONWARNINGHANDLER.fb ---- *)
FUNCTION_BLOCK L_UBUP_CONDITIONWARNINGHANDLER
VAR_INPUT
	ITFREQUEST : L_UBUP_IRequest;
END_VAR
VAR_OUTPUT
	XCONDITIONERROR : BOOL;
	EERRORIDPROPOSED : L_IE1P_Error;
END_VAR
VAR
	_ITFREQUESTACTUAL : L_UBUP_IRequest;
	_ITFSTATESERVER : L_UBUP_IStateServer;
END_VAR
END_FUNCTION_BLOCK

METHOD FB_INIT : BOOL
VAR_INPUT
	BINITRETAINS : BOOL;
	BINCOPYCODE : BOOL;
	ITFSTATESERVER : L_UBUP_IStateServer;
END_VAR
END_METHOD

METHOD RAISEWARNING
END_METHOD

METHOD RESET
END_METHOD

(* ---- L_UBUP_CRITICALSECTION.fb ---- *)
FUNCTION_BLOCK L_UBUP_CRITICALSECTION
VAR
	ISLOCKED : DWORD;
END_VAR
END_FUNCTION_BLOCK

METHOD LOCK : BOOL
END_METHOD

METHOD LOCKSTATE : BOOL
END_METHOD

METHOD REQUESTINTERFACE : BOOL
VAR_INPUT
	ID : DINT;
	PITFUNKNOWN : POINTER TO L_UBUP_IUnknown;
END_VAR
END_METHOD

METHOD UNLOCK : BOOL
END_METHOD

(* ---- L_UBUP_CYCLICCALLER.fb ---- *)
FUNCTION_BLOCK L_UBUP_CYCLICCALLER
VAR_INPUT
	HTASK : RTS_IEC_HANDLE := 0;
END_VAR
VAR
	_ITFARI : L_UBUP_IAfterReadInputs;
	_HEVENTARI : RTS_IEC_HANDLE := SysTypes.RTS_INVALID_HANDLE;
	_HINTERFACEARI : RTS_IEC_HANDLE := SysTypes.RTS_INVALID_HANDLE;
	_ITFAWO : L_UBUP_IAfterWriteOutputs;
	_HEVENTAWO : RTS_IEC_HANDLE := SysTypes.RTS_INVALID_HANDLE;
	_HINTERFACEAWO : RTS_IEC_HANDLE := SysTypes.RTS_INVALID_HANDLE;
	_ITFBRI : L_UBUP_IBeforeReadInputs;
	_HEVENTBRI : RTS_IEC_HANDLE := SysTypes.RTS_INVALID_HANDLE;
	_HINTERFACEBRI : RTS_IEC_HANDLE := SysTypes.RTS_INVALID_HANDLE;
	_ITFBWO : L_UBUP_IBeforeWriteOutputs;
	_HEVENTBWO : RTS_IEC_HANDLE := SysTypes.RTS_INVALID_HANDLE;
	_HINTERFACEBWO : RTS_IEC_HANDLE := SysTypes.RTS_INVALID_HANDLE;
	_ITFRIE : L_UBUP_IReadInputsExit;
	_HEVENTRIE : RTS_IEC_HANDLE := SysTypes.RTS_INVALID_HANDLE;
	_HINTERFACERIE : RTS_IEC_HANDLE := SysTypes.RTS_INVALID_HANDLE;
	_ITFWOE : L_UBUP_IWriteOutputsEntry;
	_HEVENTWOE : RTS_IEC_HANDLE := SysTypes.RTS_INVALID_HANDLE;
	_HINTERFACEWOE : RTS_IEC_HANDLE := SysTypes.RTS_INVALID_HANDLE;
	_ITFAIE : L_UBUP_IAfterReadInputsExit;
	_HEVENTAIE : RTS_IEC_HANDLE := SysTypes.RTS_INVALID_HANDLE;
	_HINTERFACEAIE : RTS_IEC_HANDLE := SysTypes.RTS_INVALID_HANDLE;
	_ITFAOE : L_UBUP_IAfterWriteOutputsExit;
	_HEVENTAOE : RTS_IEC_HANDLE := SysTypes.RTS_INVALID_HANDLE;
	_HINTERFACEAOE : RTS_IEC_HANDLE := SysTypes.RTS_INVALID_HANDLE;
	_ITFBIE : L_UBUP_IBeforeReadInputsEntry;
	_HEVENTBIE : RTS_IEC_HANDLE := SysTypes.RTS_INVALID_HANDLE;
	_HINTERFACEBIE : RTS_IEC_HANDLE := SysTypes.RTS_INVALID_HANDLE;
	_ITFBOE : L_UBUP_IBeforeWriteOutputsEntry;
	_HEVENTBOE : RTS_IEC_HANDLE := SysTypes.RTS_INVALID_HANDLE;
	_HINTERFACEBOE : RTS_IEC_HANDLE := SysTypes.RTS_INVALID_HANDLE;
	_ITFBRP : L_UBUP_IBreakpoint;
	_HEVENTBRP : RTS_IEC_HANDLE := SysTypes.RTS_INVALID_HANDLE;
	_HINTERFACEBRP : RTS_IEC_HANDLE := SysTypes.RTS_INVALID_HANDLE;
	_ITFEXC : L_UBUP_IException;
	_HEVENTEXC : RTS_IEC_HANDLE := SysTypes.RTS_INVALID_HANDLE;
	_HINTERFACEEXC : RTS_IEC_HANDLE := SysTypes.RTS_INVALID_HANDLE;
	_ITASKINDEX : INT;
	_HTASK : RTS_IEC_HANDLE;
	_PSCSYSTASKINFO : POINTER TO SYS_TASK_INFO;
	_UDIOSPRIORITY : UDINT;
	_UDIPRIORITY : UDINT;
	_UDITASKINTERVAL : UDINT;
	_HTASKBUS : RTS_IEC_HANDLE;
	_UDIPRIORITYBUS : UDINT;
	_XAPPISRUNNING : BOOL;
	_CAPPSTATERUN : UDINT := 1;
	_CAPPSTATESTOP : UDINT := 2;
END_VAR
END_FUNCTION_BLOCK

METHOD EVENTCALLBACK : SysTypes.RTS_IEC_RESULT
VAR_INPUT
	PEVENTPARAM : POINTER TO EventParam;
END_VAR
END_METHOD

METHOD FB_EXIT : BOOL
VAR_INPUT
	BINCOPYCODE : BOOL;
END_VAR
END_METHOD

METHOD FB_INIT : BOOL
VAR_INPUT
	BINITRETAINS : BOOL;
	BINCOPYCODE : BOOL;
	ITFCLIENT : __SYSTEM.IQueryInterface;
END_VAR
END_METHOD

METHOD FB_REINIT : BOOL
END_METHOD

METHOD REGISTEREVENTS
END_METHOD

METHOD UNREGISTEREVENTS
END_METHOD

(* ---- L_UBUP_DOUBLELINKEDLISTCONTROL.fb ---- *)
FUNCTION_BLOCK L_UBUP_DOUBLELINKEDLISTCONTROL
VAR
	_PANODES : POINTER TO ARRAY [1..16#FFFFF] OF L_UBUP_ListNode;
	_DWNODESCOUNT : DWORD;
	_DWELMCOUNT : DWORD;
	_DWFIRST : DWORD;
	_DWLAST : DWORD;
	_XLISTISEMPTY : BOOL := TRUE;
	_XLISTISFULL : BOOL := FALSE;
	_DWCURRENT : DWORD;
	CAPACITY : DWORD;
	COUNT : DWORD;
	CURRENT : DWORD;
	FIRSTARRIDX : DWORD;
	HASNEXT : BOOL;
	HASPREV : BOOL;
	ISEMPTY : BOOL;
	ISFULL : BOOL;
	LASTARRIDX : DWORD;
END_VAR
END_FUNCTION_BLOCK

METHOD NEXT : DWORD
END_METHOD

METHOD PREV : DWORD
END_METHOD

METHOD REWIND
VAR_OUTPUT
	DWARRAYIDXSTART : DWORD;
END_VAR
END_METHOD

METHOD APPEND : BOOL
VAR_OUTPUT
	DWARRIDX : DWORD;
END_VAR
END_METHOD

METHOD GETARRIDXOF : DWORD
VAR_INPUT
	DWPOSITION : DWORD;
END_VAR
END_METHOD

METHOD GETMAX : DWORD
VAR_INPUT
	ITFCOMPARER : L_UBUP_IComparer;
END_VAR
END_METHOD

METHOD GETPOSITIONOF : DWORD
VAR_INPUT
	DWARRIDX : DWORD;
END_VAR
END_METHOD

METHOD INSERTAFTER : BOOL
VAR_INPUT
	DWARRIDX : DWORD;
END_VAR
VAR_OUTPUT
	DWNEXTIDX : DWORD;
END_VAR
END_METHOD

METHOD INSERTBEFORE : BOOL
VAR_INPUT
	DWARRIDX : DWORD;
END_VAR
VAR_OUTPUT
	DWPREVIDX : DWORD;
END_VAR
END_METHOD

METHOD PREPEND : BOOL
VAR_OUTPUT
	DWARRIDX : DWORD;
END_VAR
END_METHOD

METHOD REMOVE : BOOL
VAR_INPUT
	DWARRIDX : DWORD;
END_VAR
END_METHOD

METHOD SHIFTNEXT : BOOL
VAR_INPUT
	DWARRIDX : DWORD;
END_VAR
END_METHOD

METHOD SHIFTPREV : BOOL
VAR_INPUT
	DWARRIDX : DWORD;
END_VAR
END_METHOD

METHOD SORT : BOOL
VAR_INPUT
	ITFCOMPARER : L_UBUP_IComparer;
END_VAR
END_METHOD

METHOD SWAP : BOOL
VAR_INPUT
	DWARRIDX1 : DWORD;
	DWARRIDX2 : DWORD;
END_VAR
END_METHOD

METHOD TRYAPPEND : BOOL
VAR_INPUT
	DWARRIDX : DWORD;
END_VAR
END_METHOD

METHOD TRYPREPEND : BOOL
VAR_INPUT
	DWARRIDX : DWORD;
END_VAR
END_METHOD

METHOD EVALMEMORYPROVIDER
VAR_INPUT
	ITFMEMORYPROVIDER : L_UBUP_IMemoryProvider;
END_VAR
END_METHOD

METHOD REQUESTINTERFACE : BOOL
VAR_INPUT
	ID : DINT;
	PITFUNKNOWN : POINTER TO L_UBUP_IUnknown;
END_VAR
END_METHOD

METHOD FB_INIT : BOOL
VAR_INPUT
	BINITRETAINS : BOOL;
	BINCOPYCODE : BOOL;
	ITFNODES : L_UBUP_IMemoryProvider;
END_VAR
END_METHOD

METHOD FREEARRIDX : DWORD
END_METHOD

METHOD ISFREE : BOOL
VAR_INPUT
	DWARRIDX : DWORD;
END_VAR
END_METHOD

METHOD SETFIRST
VAR_INPUT
	DWARRIDX : DWORD;
END_VAR
END_METHOD

(* ---- L_UBUP_DOUBLELINKEDLISTNODES.fb ---- *)
FUNCTION_BLOCK L_UBUP_DOUBLELINKEDLISTNODES EXTENDS L_UBUP_DoubleLinkedListNodes100Cnt
END_FUNCTION_BLOCK

(* ---- L_UBUP_DOUBLELINKEDLISTNODES1000CNT.fb ---- *)
FUNCTION_BLOCK L_UBUP_DOUBLELINKEDLISTNODES1000CNT EXTENDS L_UBUP_MemoryProvider
VAR
	ADOUBLELINKEDLISTNODES : ARRAY [1..1000] OF L_UBUP_ListNode;
	PTR : POINTER TO BYTE;
	SIZE : UDINT;
END_VAR
END_FUNCTION_BLOCK

(* ---- L_UBUP_DOUBLELINKEDLISTNODES100CNT.fb ---- *)
FUNCTION_BLOCK L_UBUP_DOUBLELINKEDLISTNODES100CNT EXTENDS L_UBUP_MemoryProvider
VAR
	ADOUBLELINKEDLISTNODES : ARRAY [1..100] OF L_UBUP_ListNode;
	PTR : POINTER TO BYTE;
	SIZE : UDINT;
END_VAR
END_FUNCTION_BLOCK

(* ---- L_UBUP_DOUBLELINKEDLISTNODES5CNT.fb ---- *)
FUNCTION_BLOCK L_UBUP_DOUBLELINKEDLISTNODES5CNT EXTENDS L_UBUP_MemoryProvider
VAR
	ADOUBLELINKEDLISTNODES : ARRAY [1..5] OF L_UBUP_ListNode;
	PTR : POINTER TO BYTE;
	SIZE : UDINT;
END_VAR
END_FUNCTION_BLOCK

(* ---- L_UBUP_DURATION.fb ---- *)
FUNCTION_BLOCK L_UBUP_DURATION
VAR_OUTPUT
	STARTTIME : SYSTIME;
	STOPTIME : SYSTIME;
	DURATION : SYSTIME;
END_VAR
END_FUNCTION_BLOCK

METHOD START
END_METHOD

METHOD STOP
END_METHOD

(* ---- L_UBUP_DYNMEMORYPROVIDER.fb ---- *)
FUNCTION_BLOCK L_UBUP_DYNMEMORYPROVIDER EXTENDS L_UBUP_MemoryProvider
VAR
	_PMEM : POINTER TO ARRAY [1..16#FFFF] OF BYTE;
	_DWMEMSIZE : DWORD;
	PTR : POINTER TO BYTE;
	SIZE : UDINT;
END_VAR
END_FUNCTION_BLOCK

METHOD FB_EXIT : BOOL
VAR_INPUT
	BINCOPYCODE : BOOL;
END_VAR
END_METHOD

METHOD FB_INIT : BOOL
VAR_INPUT
	BINITRETAINS : BOOL;
	BINCOPYCODE : BOOL;
	DWMEMSIZE : DWORD;
END_VAR
END_METHOD

(* ---- L_UBUP_FBCONTAINER.fb ---- *)
FUNCTION_BLOCK L_UBUP_FBCONTAINER EXTENDS InstanceBase
VAR
	_ITFOWNER : L_UBUP_IFBPool;
	_XWHANDLE : __XWORD;
	_XOCCUPIED : BOOL;
	CLASSID : DINT;
	INSTANCEPTR : POINTER TO BYTE;
	OBJECTID : DWORD;
	OCCUPIED : BOOL;
	PRVINSTFACTORY : FBF.IFactory;
	PRVNEXTINST : FBF.IInstance;
	PRVPREVINST : FBF.IInstance;
END_VAR
END_FUNCTION_BLOCK

METHOD DISPOSE : BOOL
END_METHOD

METHOD PRVINSTINIT : FBF.ERROR
VAR_INPUT
	ITFDATA : FBF.IData;
END_VAR
END_METHOD

METHOD PRVINSTRELEASE : BOOL
END_METHOD

METHOD PRVINSTRETAIN : BOOL
END_METHOD

METHOD FREE : BOOL
END_METHOD

METHOD OCCUPY : BOOL
VAR_INPUT
	ITFOWNER : L_UBUP_IFBPool;
	XWHANDLE : __XWORD;
END_VAR
END_METHOD

METHOD REQUESTINTERFACE : BOOL
VAR_INPUT
	ID : DINT;
	PITFUNKNOWN : POINTER TO L_UBUP_IUnknown;
END_VAR
END_METHOD

(* ---- L_UBUP_FBPOOL.fb ---- *)
FUNCTION_BLOCK L_UBUP_FBPOOL
VAR
	USEGLOBAL : BOOL;
END_VAR
END_FUNCTION_BLOCK

METHOD FREEINSTANCE : BOOL
VAR_INPUT
	ITFINSTANCE : L_UBUP_IPoolInstance;
	XWHANDLE : __XWORD;
END_VAR
END_METHOD

METHOD GETCAPACITY : BOOL
VAR_INPUT
	ECLASSID : DINT;
END_VAR
VAR_OUTPUT
	DWCAPACITY : DWORD;
END_VAR
END_METHOD

METHOD QUERYINSTANCE : BOOL
VAR_INPUT
	ECLASSID : DINT;
END_VAR
VAR_IN_OUT
	ITFINSTANCE : L_UBUP_IPoolInstance;
END_VAR
END_METHOD

METHOD FB_INIT : BOOL
VAR_INPUT
	BINITRETAINS : BOOL;
	BINCOPYCODE : BOOL;
END_VAR
END_METHOD

METHOD FB_AFTERGLOBALINIT : BOOL
END_METHOD

METHOD FREERESOURCE
END_METHOD

METHOD GETFB : L_UBUP_IPoolInstance
VAR_INPUT
	ECLASSID : DINT;
	DWARRIDX : DWORD;
END_VAR
END_METHOD

METHOD GETFBCONTROL : L_UBUP_IListControl
VAR_INPUT
	ECLASSID : DINT;
END_VAR
END_METHOD

METHOD OCCUPYRESOURCE : BOOL
VAR_INPUT
	ECLASSID : DINT;
END_VAR
END_METHOD

METHOD SETCAPACITY
VAR_INPUT
	ITFLISTCONTROL : L_UBUP_IListControl;
	DWCAPACITY : DWORD;
END_VAR
END_METHOD

METHOD SETCAPACITYALL
END_METHOD

(* ---- L_UBUP_FBPOOLCOLLECTION.fb ---- *)
FUNCTION_BLOCK L_UBUP_FBPOOLCOLLECTION
VAR
	_AITFFBPOOL : ARRAY [1..c_dwMaxPools] OF L_UBUP_IFBPool;
	C_DWMAXPOOLS : DWORD := 10;
END_VAR
END_FUNCTION_BLOCK

METHOD REGISTERPOOL : BOOL
VAR_INPUT
	ITFFBPOOL : L_UBUP_IFBPool;
END_VAR
END_METHOD

METHOD FREEINSTANCE : BOOL
VAR_INPUT
	ITFINSTANCE : L_UBUP_IPoolInstance;
	XWHANDLE : __XWORD;
END_VAR
END_METHOD

METHOD GETCAPACITY : BOOL
VAR_INPUT
	ECLASSID : DINT;
END_VAR
VAR_OUTPUT
	DWCAPACITY : DWORD;
END_VAR
END_METHOD

METHOD QUERYINSTANCE : BOOL
VAR_INPUT
	ECLASSID : DINT;
END_VAR
VAR_IN_OUT
	ITFINSTANCE : L_UBUP_IPoolInstance;
END_VAR
END_METHOD

(* ---- L_UBUP_FBPOOLFACTORY.fb ---- *)
FUNCTION_BLOCK L_UBUP_FBPOOLFACTORY EXTENDS FactoryBase
VAR
	_AITFINSTANCE : ARRAY [1..100] OF L_UBUP_IPoolInstance;
	_FBCONTROLNODES : L_UBUP_DoubleLinkedListNodes100Cnt;
	_FBCONTROL : L_UBUP_DoubleLinkedListControl;
	_ECLASSID : DINT;
	_XFIRSTCALL : BOOL := TRUE;
	_PPOOLADR : POINTER TO BYTE;
	_DWPOOLSIZE : DWORD;
	INSTSIZE : DWORD;
	PRVINSTCOUNT : CAA.COUNT;
	PRVINSTPOOLADR : CAA.PVOID;
	PRVINSTPOOLEXTENDSFACTOR : USINT;
	PRVINSTPOOLSIZE : CAA.SIZE;
	PRVINSTSIZE : CAA.SIZE;
END_VAR
END_FUNCTION_BLOCK

METHOD CREATEPOOL
VAR_INPUT
	ECLASSID : DINT;
END_VAR
END_METHOD

METHOD PRVALLOCINSTMEM : CAA.HANDLE
VAR_OUTPUT
	EERROR : FBF.ERROR;
END_VAR
END_METHOD

METHOD PRVFREEINSTMEM : BOOL
VAR_INPUT
	HINST : CAA.HANDLE;
END_VAR
END_METHOD

METHOD PRVGETINSTPOINTER : CAA.PVOID
VAR_INPUT
	HINST : CAA.HANDLE;
END_VAR
END_METHOD

METHOD PRVINSERTINST : BOOL
VAR_INPUT
	ITFINST : FBF.IInstance;
END_VAR
END_METHOD

METHOD PRVINSTINIT : BOOL
VAR_INPUT
	ITFINST : FBF.IInstance;
	HINST : CAA.HANDLE;
	ITFDATA : FBF.IData;
END_VAR
VAR_OUTPUT
	EERROR : FBF.ERROR;
END_VAR
END_METHOD

METHOD PRVREMOVEINST : BOOL
VAR_INPUT
	ITFINST : FBF.IInstance;
END_VAR
END_METHOD

METHOD FREEINSTANCE : BOOL
VAR_INPUT
	ITFINSTANCE : L_UBUP_IPoolInstance;
	XWHANDLE : __XWORD;
END_VAR
END_METHOD

METHOD GETCAPACITY : BOOL
VAR_INPUT
	ECLASSID : DINT;
END_VAR
VAR_OUTPUT
	DWCAPACITY : DWORD;
END_VAR
END_METHOD

METHOD QUERYINSTANCE : BOOL
VAR_INPUT
	ECLASSID : DINT;
END_VAR
VAR_IN_OUT
	ITFINSTANCE : L_UBUP_IPoolInstance;
END_VAR
END_METHOD

METHOD EVALMEMORYPROVIDER
VAR_INPUT
	ITFMEMORYPROVIDER : L_UBUP_IMemoryProvider;
END_VAR
END_METHOD

METHOD FB_INIT : BOOL
VAR_INPUT
	BINITRETAINS : BOOL;
	BINCOPYCODE : BOOL;
	ITFMEMORY : L_UBUP_IMemoryProvider;
END_VAR
END_METHOD

METHOD CREATEINST : BOOL
VAR_INPUT
	ECLASSID : DINT;
END_VAR
VAR_IN_OUT
	ITFINSTANCE : L_UBUP_IPoolInstance;
END_VAR
END_METHOD

(* ---- L_UBUP_FREERUNTASK.fb ---- *)
FUNCTION_BLOCK L_UBUP_FREERUNTASK
VAR_INPUT
	XEXECUTE : BOOL;
	EFREERUNTASKTYPE : L_UBUP_FreeRunTaskType;
END_VAR
VAR_OUTPUT
	XBUSY : BOOL;
	XDONE : BOOL;
	XERROR : BOOL;
	EERRORID : L_IE1P_Error;
	XFREERUNTASKBUSY : BOOL;
	DURATION : SYSTIME;
END_VAR
VAR
	UDIRESULT : UDINT;
	EFREERUNTASKTYPEACTUAL : L_UBUP_FreeRunTaskType;
	_MODEL : L_UBUP_BehaviourModel_ETrig;
END_VAR
END_FUNCTION_BLOCK

METHOD CYCLICACTION
VAR_INPUT
	ITFTIMINGCONTROLLER : L_UBUP_ITimingController;
END_VAR
VAR_OUTPUT
	XCOMPLETE : BOOL;
	XABORT : BOOL;
	IERRORID : INT;
END_VAR
END_METHOD

METHOD FINALIZEACTION
VAR_INPUT
	XABORTPROPOSED : BOOL;
	IERRORIDPROPOSED : INT;
END_VAR
VAR_OUTPUT
	XCOMPLETE : BOOL;
	XABORT : BOOL;
	IERRORID : INT;
END_VAR
END_METHOD

METHOD RESETACTION
VAR_OUTPUT
	XCOMPLETE : BOOL;
END_VAR
END_METHOD

METHOD STARTACTION
VAR_OUTPUT
	XCOMPLETE : BOOL;
	IERRORID : INT;
END_VAR
END_METHOD

METHOD FB_INIT : BOOL
VAR_INPUT
	BINITRETAINS : BOOL;
	BINCOPYCODE : BOOL;
END_VAR
END_METHOD

METHOD ABORT : UDINT
END_METHOD

METHOD EXECUTE : UDINT
END_METHOD

METHOD CUSTOMIZEERRORCODE : L_IE1P_Error
VAR_INPUT
	IERRORID : INT;
END_VAR
END_METHOD

METHOD EXECUTEIMPL : UDINT
END_METHOD

METHOD EXTERNALFREERUNTASK
END_METHOD

(* ---- L_UBUP_HISTOGRAM.fb ---- *)
FUNCTION_BLOCK L_UBUP_HISTOGRAM
VAR_INPUT
	XENABLE : BOOL;
	XRESET : BOOL;
	LRNEXT : LREAL;
END_VAR
VAR_OUTPUT
	XBUSY : BOOL;
	XERROR : BOOL;
	EERRORID : L_IE1P_Error;
END_VAR
VAR
	_PLIHISTO : POINTER TO LINT;
	_DWHISTODATASIZE : DWORD;
	_DWHISTOELMS : DWORD;
	_LRHISTOSTART : LREAL;
	_LRRESOLUTION : LREAL;
	_LRHISTOSTOP : LREAL;
	_ITFHISTOMEM : L_UBUP_IMemoryProvider;
	_MODEL : L_UBUP_BehaviourModel_LConC;
END_VAR
END_FUNCTION_BLOCK

METHOD CYCLICACTION
VAR_INPUT
	ITFTIMINGCONTROLLER : L_UBUP_ITimingController;
END_VAR
VAR_OUTPUT
	XCOMPLETE : BOOL;
	XABORT : BOOL;
	IERRORID : INT;
END_VAR
END_METHOD

METHOD FINALIZEACTION
VAR_INPUT
	XABORTPROPOSED : BOOL;
	IERRORIDPROPOSED : INT;
END_VAR
VAR_OUTPUT
	XCOMPLETE : BOOL;
	XABORT : BOOL;
	IERRORID : INT;
END_VAR
END_METHOD

METHOD RESETACTION
VAR_OUTPUT
	XCOMPLETE : BOOL;
END_VAR
END_METHOD

METHOD STARTACTION
VAR_OUTPUT
	XCOMPLETE : BOOL;
	IERRORID : INT;
END_VAR
END_METHOD

METHOD EVALMEMORYPROVIDER
VAR_INPUT
	ITFMEMORYPROVIDER : L_UBUP_IMemoryProvider;
END_VAR
END_METHOD

METHOD FB_INIT : BOOL
VAR_INPUT
	BINITRETAINS : BOOL;
	BINCOPYCODE : BOOL;
	LRRESOLUTION : LREAL;
	LRHISTOSTART : LREAL;
	ITFHISTOMEM : L_UBUP_IMemoryProvider;
END_VAR
END_METHOD

METHOD RESET
END_METHOD

(* ---- L_UBUP_HISTOGRAMSTATESERVER.fb ---- *)
FUNCTION_BLOCK L_UBUP_HISTOGRAMSTATESERVER
VAR_INPUT
	XENABLE : BOOL;
	XRESET : BOOL;
END_VAR
VAR_OUTPUT
	XBUSY : BOOL;
	PHISTO_1 : POINTER TO ARRAY [1..100] OF LINT;
	PHISTO_2 : POINTER TO ARRAY [1..100] OF LINT;
	PHISTO_3 : POINTER TO ARRAY [1..100] OF LINT;
	PHISTO_4 : POINTER TO ARRAY [1..100] OF LINT;
	PHISTO_5 : POINTER TO ARRAY [1..100] OF LINT;
	PHISTO_6 : POINTER TO ARRAY [1..100] OF LINT;
	PHISTO_7 : POINTER TO ARRAY [1..100] OF LINT;
	PHISTO_8 : POINTER TO ARRAY [1..100] OF LINT;
	PHISTO_9 : POINTER TO ARRAY [1..100] OF LINT;
	PHISTO_10 : POINTER TO ARRAY [1..100] OF LINT;
	PHISTO_11 : POINTER TO ARRAY [1..100] OF LINT;
	PHISTO_12 : POINTER TO ARRAY [1..100] OF LINT;
	PHISTO_13 : POINTER TO ARRAY [1..100] OF LINT;
	PHISTO_14 : POINTER TO ARRAY [1..100] OF LINT;
	PHISTO_15 : POINTER TO ARRAY [1..100] OF LINT;
	PHISTO_16 : POINTER TO ARRAY [1..100] OF LINT;
	PHISTO_17 : POINTER TO ARRAY [1..100] OF LINT;
END_VAR
VAR_IN_OUT
	ATIMESTAMP : ARRAY [1..17] OF SYSTIME;
END_VAR
VAR
	_AHISTODATA : ARRAY [1..17] OF L_UBUP_MemoryProvider100LINT;
	_PAHISTO : ARRAY [1..17] OF POINTER TO L_UBUP_Histogram;
	_HISTO_1 : L_UBUP_Histogram;
	_HISTO_2 : L_UBUP_Histogram;
	_HISTO_3 : L_UBUP_Histogram;
	_HISTO_4 : L_UBUP_Histogram;
	_HISTO_5 : L_UBUP_Histogram;
	_HISTO_6 : L_UBUP_Histogram;
	_HISTO_7 : L_UBUP_Histogram;
	_HISTO_8 : L_UBUP_Histogram;
	_HISTO_9 : L_UBUP_Histogram;
	_HISTO_10 : L_UBUP_Histogram;
	_HISTO_11 : L_UBUP_Histogram;
	_HISTO_12 : L_UBUP_Histogram;
	_HISTO_13 : L_UBUP_Histogram;
	_HISTO_14 : L_UBUP_Histogram;
	_HISTO_15 : L_UBUP_Histogram;
	_HISTO_16 : L_UBUP_Histogram;
	_HISTO_17 : L_UBUP_Histogram;
	_MODEL : L_UBUP_BehaviourModel_LConC;
END_VAR
END_FUNCTION_BLOCK

METHOD CYCLICACTION
VAR_INPUT
	ITFTIMINGCONTROLLER : L_UBUP_ITimingController;
END_VAR
VAR_OUTPUT
	XCOMPLETE : BOOL;
	XABORT : BOOL;
	IERRORID : INT;
END_VAR
END_METHOD

METHOD FINALIZEACTION
VAR_INPUT
	XABORTPROPOSED : BOOL;
	IERRORIDPROPOSED : INT;
END_VAR
VAR_OUTPUT
	XCOMPLETE : BOOL;
	XABORT : BOOL;
	IERRORID : INT;
END_VAR
END_METHOD

METHOD RESETACTION
VAR_OUTPUT
	XCOMPLETE : BOOL;
END_VAR
END_METHOD

METHOD STARTACTION
VAR_OUTPUT
	XCOMPLETE : BOOL;
	IERRORID : INT;
END_VAR
END_METHOD

METHOD ALLOCPOINTADR
VAR_OUTPUT
	IERRORID : INT;
END_VAR
END_METHOD

(* ---- L_UBUP_INSTANCE.fb ---- *)
FUNCTION_BLOCK L_UBUP_INSTANCE
VAR
	_DWOBJID : DWORD;
	CLASSID : DINT;
	OBJECTID : DWORD;
END_VAR
END_FUNCTION_BLOCK

METHOD REQUESTINTERFACE : BOOL
VAR_INPUT
	ID : DINT;
	PITFUNKNOWN : POINTER TO L_UBUP_IUnknown;
END_VAR
END_METHOD

METHOD FB_INIT : BOOL
VAR_INPUT
	BINITRETAINS : BOOL;
	BINCOPYCODE : BOOL;
END_VAR
END_METHOD

(* ---- L_UBUP_JOB.fb ---- *)
FUNCTION_BLOCK L_UBUP_JOB EXTENDS L_UBUP_PoolInstance
VAR
	_EERRORID : L_IE1P_Error;
	_XABORT : BOOL;
	_XDONE : BOOL;
	_ITFSENDER : L_UBUP_ICommand;
	_ITFREPORT : L_UBUP_IJobReport;
	_ITFPREVJOB : L_UBUP_IJob;
	_ITFNEXTJOB : L_UBUP_IJob;
	_DWCALLID : DWORD := L_UBUP_Internal.g_dwCallIDUnassigned;
	_ECMDID : L_UBUP_ClassID;
	_ESTATE : L_UBUP_JobState;
	_CLIENTPROXY : L_UBUP_StateClientProxy;
	_STATESERVER : L_UBUP_StateServer;
	_DWARRIDX : DWORD;
	_DIREFCOUNTER : DINT;
	_SINSTANCESTR : STRING;
	FB_TRANSITION2ERROR : L_UBUP_RequestTransitionEdge;
	FB_TRANSITION2PENDINGFORWORKING : L_UBUP_RequestTransitionEdge;
	FB_TRANSITION2WORKING : L_UBUP_RequestTransitionEdge;
	FB_TRANSITION2PENDINGFORFINISH : L_UBUP_RequestTransitionEdge;
	FB_TRANSITION2READYFORRELEASE : L_UBUP_RequestTransitionEdge;
	FB_TRANSITION2PREPARERELEASE : L_UBUP_RequestTransitionEdge;
	BLOCKNEXT : BOOL;
	CALLID : DWORD;
	CANCELFINISHNEXT : BOOL;
	CLASSID : DINT;
	CMDID : L_UBUP_ClassID;
	ISAPPEND : BOOL;
	ISBLOCKED : BOOL;
	ISLINKED : BOOL;
	ISREADYFORRELEASE : BOOL;
	ITFCATEGORY : L_UBUP_ICategory;
	ITFJOBACTION : L_UBUP_IJobAction;
	ITFMAPSTATE : L_UBUP_IMapState;
	JOBSTATE : L_UBUP_JobState;
	MAPPRIO : INT;
	MAPSTATE : INT;
	NEXT : L_UBUP_IJob;
	PREV : L_UBUP_IJob;
	REJECTIFABORTED : BOOL;
	REJECTIFPENDING : BOOL;
END_VAR
END_FUNCTION_BLOCK

METHOD CLASSIFY : BOOL
VAR_INPUT
	ECATEGORY : DINT;
END_VAR
END_METHOD

METHOD EXPAND : BOOL
VAR_INPUT
	ITFSENDER : L_UBUP_ICommand;
	DWCALLID : DWORD;
END_VAR
VAR_OUTPUT
	EERRORID : L_IE1P_Error;
END_VAR
END_METHOD

METHOD HANDOVERRESOURCE : BOOL
VAR_INPUT
	ITFRESOURCE : L_UBUP_IUnknown;
END_VAR
END_METHOD

METHOD LINK : BOOL
VAR_INPUT
	ITFJOB : L_UBUP_IJob;
	XPREV : BOOL;
END_VAR
VAR_OUTPUT
	EERRORID : L_IE1P_Error;
END_VAR
END_METHOD

METHOD RELEASE
END_METHOD

METHOD ABORT
END_METHOD

METHOD CYCLE
VAR_OUTPUT
	ESTATE : L_UBUP_JobState;
	EERRORID : L_IE1P_Error;
END_VAR
END_METHOD

METHOD FINISH
END_METHOD

METHOD UPDATEREPORTDATA : BOOL
VAR_INPUT
	DWCALLID : DWORD;
END_VAR
VAR_IN_OUT
	SCREPORT : L_UBUP_ReportData;
END_VAR
END_METHOD

METHOD UPDATEREPORTRECEIVER : BOOL
VAR_INPUT
	ITFJOBREPORT : L_UBUP_IJobReport;
END_VAR
END_METHOD

METHOD GET_EERRORID : L_IE1P_Error
END_METHOD

METHOD GET_XACTIVE : BOOL
END_METHOD

METHOD GET_XBUSY : BOOL
END_METHOD

METHOD GET_XCOMMANDABORTED : BOOL
END_METHOD

METHOD GET_XDONE : BOOL
END_METHOD

METHOD GET_XINITIAL : BOOL
END_METHOD

METHOD DECCOUNTER : DINT
END_METHOD

METHOD INCCOUNTER : DINT
END_METHOD

METHOD CALLFBS
VAR_INPUT
	ECASE : L_UBUP_StateHandleCase;
END_VAR
END_METHOD

METHOD CALLSTATE
VAR_INPUT
	ITFSTATESERVER : L_UBUP_IStateServer;
	ISTATE : INT;
	ECASE : L_UBUP_StateHandleCase;
END_VAR
END_METHOD

METHOD CHECKTRANSITION
VAR_INPUT
	ITFSTATESERVER : L_UBUP_IStateServer;
END_VAR
END_METHOD

METHOD DISABLECLIENT : BOOL
VAR_INPUT
	XFIRSTCALL : BOOL;
END_VAR
END_METHOD

METHOD ENABLECLIENT : BOOL
VAR_INPUT
	XFIRSTCALL : BOOL;
END_VAR
END_METHOD

METHOD FINALIZECYCLE
END_METHOD

METHOD LEAVESTATE
END_METHOD

METHOD PREPARECYCLE
END_METHOD

METHOD PREPARESTATECHANGE
END_METHOD

METHOD STIMULATETRANSITION
VAR_INPUT
	ECASE : L_UBUP_StateHandleCase;
END_VAR
END_METHOD

METHOD UPDATECONDITIONERROR : BOOL
VAR_INPUT
	ITFREQUEST : L_UBUP_IRequest;
END_VAR
END_METHOD

METHOD REQUESTINTERFACE : BOOL
VAR_INPUT
	ID : DINT;
	PITFUNKNOWN : POINTER TO L_UBUP_IUnknown;
END_VAR
END_METHOD

METHOD CALLERRORHANDLER
VAR_INPUT
	EERRORID : L_IE1P_Error;
END_VAR
END_METHOD

METHOD STATE_ERROR
VAR_INPUT
	ECASE : L_UBUP_StateHandleCase;
	ITFSTATESERVER : L_UBUP_IStateServer;
END_VAR
END_METHOD

METHOD STATE_PENDINGFORFINISH
VAR_INPUT
	ECASE : L_UBUP_StateHandleCase;
	ITFSTATESERVER : L_UBUP_IStateServer;
END_VAR
END_METHOD

METHOD STATE_PENDINGFORWORKING
VAR_INPUT
	ECASE : L_UBUP_StateHandleCase;
	ITFSTATESERVER : L_UBUP_IStateServer;
END_VAR
END_METHOD

METHOD STATE_PREPARERELEASE
VAR_INPUT
	ECASE : L_UBUP_StateHandleCase;
	ITFSTATESERVER : L_UBUP_IStateServer;
END_VAR
END_METHOD

METHOD STATE_WORKING
VAR_INPUT
	ECASE : L_UBUP_StateHandleCase;
	ITFSTATESERVER : L_UBUP_IStateServer;
END_VAR
END_METHOD

(* ---- L_UBUP_JOBADMINSTRATION.fb ---- *)
FUNCTION_BLOCK L_UBUP_JOBADMINSTRATION EXTENDS AsyncBaseClass
VAR_OUTPUT
	XDONE : BOOL;
	XERROR : BOOL;
	WERROR : WORD;
END_VAR
VAR
	HEVENTCOMMCYCLE : RTS_IEC_HANDLE;
	HINTERFACECOMMCYCLE : RTS_IEC_HANDLE;
	ITFCALLBACK : CmpEventMgr.ICmpEventCallback;
	DWEVENTCOUNTER1 : DWORD;
	XINITALJOBADDED : BOOL;
	UDIOPERATINGSYSTEMID : UDINT;
	COUNT1 : DWORD;
	COUNT2 : DWORD;
	COUNT3 : DWORD;
	ALMDATA : ARRAY [1..c_MaxCount] OF L_UBUP_ILMData;
	AXBUSY : ARRAY [1..c_MaxJobs] OF BOOL;
	AACTIVELMDATA : ARRAY [1..c_MaxJobs] OF L_UBUP_ILMData;
	JOB : ARRAY [1..c_MaxJobs] OF RTS_IEC_HANDLE;
	JOBSTATE : ARRAY [1..c_MaxJobs] OF UDINT;
	AJOBPARA : ARRAY [1..c_MaxJobs] OF L_UBUP_LMParamCallFunction;
	FIRSTINITJOBSTATE : UDINT;
	FIRSTINITJOB : RTS_IEC_HANDLE;
	FIRSTINITJOBCALLED : BOOL;
	XINITJOBACTIVE : BOOL := TRUE;
	WINITCOUNTER : WORD;
	IDX : WORD;
	JOBCOUNT : WORD;
	WSEARCHINDEX : WORD := 0;
	WFIRSTENTRY : WORD := 1;
	WLASTENTRY : WORD := 1;
	WLISTCOUNT : WORD := 0;
	WTMPCOUNT : WORD := 333;
	AWJOBLIST : ARRAY [1..c_MaxJobs] OF WORD := [1, 2, 3, 4, 5, 6, 7, 8, 9, 10];
	JOBIDX : WORD;
	DWJOBEXECUTE : DWORD;
	DWJOBDONE : DWORD;
	DWJOBERROR : DWORD;
	RESULTASYNCADD : RTS_IEC_RESULT;
	RESULTTASK : RTS_IEC_RESULT;
	ASYNCJOBPARAM : AsyncJob_Param;
	ASYNCJOBNAME : STRING := 'ReadMotionFiles';
	JOBRES : UDINT;
	C_MAXJOBS : WORD := 10;
	C_MAXSEARCHCOUNT : WORD := 10;
	C_MAXCOUNT : WORD := 100;
END_VAR
END_FUNCTION_BLOCK

METHOD DOFIRSTINITJOB : RTS_IEC_RESULT
VAR_INPUT
	PPARAM : POINTER TO L_UBUP_LMParamCallFunction;
END_VAR
END_METHOD

METHOD DOJOB : RTS_IEC_RESULT
VAR_INPUT
	PPARAM : POINTER TO L_UBUP_LMParamCallFunction;
END_VAR
END_METHOD

METHOD FINISHJOB
VAR_INPUT
	ID : WORD;
END_VAR
END_METHOD

METHOD HANDLEINITJOB : BOOL
VAR_INPUT
	XEXITHANDLING : BOOL;
END_VAR
END_METHOD

METHOD INSERTDATA : BOOL
VAR_INPUT
	ITFLMDATA : L_UBUP_ILMData;
END_VAR
END_METHOD

METHOD FB_EXIT : BOOL
VAR_INPUT
	BINCOPYCODE : BOOL;
END_VAR
END_METHOD

METHOD FB_INIT : BOOL
VAR_INPUT
	BINITRETAINS : BOOL;
	BINCOPYCODE : BOOL;
END_VAR
END_METHOD

METHOD EVENTCALLBACK : UDINT
VAR_INPUT
	PEVENTPARAM : POINTER TO EventParam;
END_VAR
END_METHOD

METHOD REGISTEREVENT
END_METHOD

METHOD UNREGISTEREVENT
END_METHOD

(* ---- L_UBUP_JOBEXECUTER.fb ---- *)
FUNCTION_BLOCK L_UBUP_JOBEXECUTER EXTENDS L_UBUP_MemoryProvider
VAR_INPUT
	XFINISH : BOOL;
	XABORT : BOOL;
	XCLEAR : BOOL;
END_VAR
VAR
	C_DWMAXJOBSEXECUTED : DWORD := 200;
	_ALISTNODES : ARRAY [1..c_dwMaxJobsExecuted] OF L_UBUP_ListNode;
	_AJOBS : ARRAY [1..c_dwMaxJobsExecuted] OF L_UBUP_IJob;
	_JOBLISTCONTROL : L_UBUP_DoubleLinkedListControl;
	_DWARRIDX : DWORD;
	_EACTUALSTATE : L_UBUP_JobState;
	_EERRORID : L_IE1P_Error;
	_XFINISH_TRIG : R_Trig;
	_XABORT_TRIG : R_Trig;
	_XCLEAR_TRIG : R_Trig;
	_ITFJOBTEMP : L_UBUP_IJob;
	_XREMOVELAST : BOOL;
	_ITFJOBRECEIVERMONITOR : L_UBUP_IJobReceiverListener;
	ITFITERATOR : L_UBUP_IIterator;
	ITFLISTCONTROL : L_UBUP_IListControl;
	PTR : POINTER TO BYTE;
	SIZE : UDINT;
END_VAR
END_FUNCTION_BLOCK

METHOD GETJOB : BOOL
VAR_INPUT
	DWARRIDX : DWORD;
END_VAR
VAR_OUTPUT
	ITFJOB : L_UBUP_IJob;
END_VAR
END_METHOD

METHOD ANNOUNCELISTENER : BOOL
VAR_INPUT
	ITFLISTENER : L_UBUP_IJobReceiverListener;
END_VAR
END_METHOD

METHOD INSERT : BOOL
VAR_INPUT
	ITFJOB : L_UBUP_IJob;
END_VAR
END_METHOD

METHOD UNPLUGLISTENER : BOOL
VAR_INPUT
	ITFLISTENER : L_UBUP_IJobReceiverListener;
END_VAR
END_METHOD

METHOD REQUESTINTERFACE : BOOL
VAR_INPUT
	ID : DINT;
	PITFUNKNOWN : POINTER TO L_UBUP_IUnknown;
END_VAR
END_METHOD

METHOD FB_INIT : BOOL
VAR_INPUT
	BINITRETAINS : BOOL;
	BINCOPYCODE : BOOL;
END_VAR
END_METHOD

(* ---- L_UBUP_JOBLISTREADER.fb ---- *)
FUNCTION_BLOCK L_UBUP_JOBLISTREADER
VAR_INPUT
	ALRITFJOBS : POINTER TO L_UBUP_IJob;
	XENABLE : BOOL;
	ITFJOBS : L_UBUP_IList;
END_VAR
VAR_OUTPUT
	XBUSY : BOOL;
	XERROR : BOOL;
	EERRORID : L_IE1P_Error;
	DWJOBCOUNT : DWORD;
END_VAR
VAR
	_JOBMANAGER : L_UBUP_JobManager;
	_MODEL : L_UBUP_BehaviourModel_LConC;
END_VAR
END_FUNCTION_BLOCK

METHOD CYCLICACTION
VAR_INPUT
	ITFTIMINGCONTROLLER : L_UBUP_ITimingController;
END_VAR
VAR_OUTPUT
	XCOMPLETE : BOOL;
	XABORT : BOOL;
	IERRORID : INT;
END_VAR
END_METHOD

METHOD FINALIZEACTION
VAR_INPUT
	XABORTPROPOSED : BOOL;
	IERRORIDPROPOSED : INT;
END_VAR
VAR_OUTPUT
	XCOMPLETE : BOOL;
	XABORT : BOOL;
	IERRORID : INT;
END_VAR
END_METHOD

METHOD RESETACTION
VAR_OUTPUT
	XCOMPLETE : BOOL;
END_VAR
END_METHOD

METHOD STARTACTION
VAR_OUTPUT
	XCOMPLETE : BOOL;
	IERRORID : INT;
END_VAR
END_METHOD

(* ---- L_UBUP_JOBMANAGER.fb ---- *)
FUNCTION_BLOCK L_UBUP_JOBMANAGER
VAR_INPUT
	XENABLE : BOOL;
	DWJOBNO : DWORD := 1;
	ITFJOBS : L_UBUP_IList;
END_VAR
VAR_OUTPUT
	XBUSY : BOOL;
	XERROR : BOOL;
	EERRORID : L_IE1P_Error;
	DWJOBCOUNT : DWORD;
	DWCALLID : DWORD := L_UBUP_Internal.g_dwCallIDUnassigned;
	EACTUALSTATE : L_UBUP_JobState;
	ITFJOB : L_UBUP_IJob;
	ECLASSID : DINT;
END_VAR
VAR
	_ITFJOBCOLLECTION : L_UBUP_IJobCollection;
	_ITFLISTCONTROL : L_UBUP_IListControl;
	_MODEL : L_UBUP_BehaviourModel_LConC;
END_VAR
END_FUNCTION_BLOCK

METHOD CYCLICACTION
VAR_INPUT
	ITFTIMINGCONTROLLER : L_UBUP_ITimingController;
END_VAR
VAR_OUTPUT
	XCOMPLETE : BOOL;
	XABORT : BOOL;
	IERRORID : INT;
END_VAR
END_METHOD

METHOD FINALIZEACTION
VAR_INPUT
	XABORTPROPOSED : BOOL;
	IERRORIDPROPOSED : INT;
END_VAR
VAR_OUTPUT
	XCOMPLETE : BOOL;
	XABORT : BOOL;
	IERRORID : INT;
END_VAR
END_METHOD

METHOD RESETACTION
VAR_OUTPUT
	XCOMPLETE : BOOL;
END_VAR
END_METHOD

METHOD STARTACTION
VAR_OUTPUT
	XCOMPLETE : BOOL;
	IERRORID : INT;
END_VAR
END_METHOD

(* ---- L_UBUP_JOBPOOLQUEUE.fb ---- *)
FUNCTION_BLOCK L_UBUP_JOBPOOLQUEUE
VAR
	C_DWCAPACITY : DWORD := 100;
	FBQUEUE : L_UBUP_QueueArrayControl;
	_ALISTENELEMENT : ARRAY [1..c_dwCapacity] OF L_UBUP_IFBPool;
END_VAR
END_FUNCTION_BLOCK

METHOD REGISTERPOOL : BOOL
VAR_INPUT
	ITFJOBPOOL : L_UBUP_IFBPool;
END_VAR
END_METHOD

METHOD GETCAPACITY : BOOL
VAR_INPUT
	ECLASSID : L_UBUP_ClassID;
END_VAR
VAR_OUTPUT
	ITFJOBPOOL : L_UBUP_IFBPool;
	DWCAPACITY : DWORD;
END_VAR
END_METHOD

METHOD QUERYINSTANCE : BOOL
VAR_INPUT
	ECLASSID : DINT;
END_VAR
VAR_OUTPUT
	ITFJOBPOOL : L_UBUP_IFBPool;
END_VAR
VAR_IN_OUT
	ITFINSTANCE : L_UBUP_IPoolInstance;
END_VAR
END_METHOD

(* ---- L_UBUP_MEMORYPROVIDER.fb ---- *)
FUNCTION_BLOCK L_UBUP_MEMORYPROVIDER
VAR
	_ITFCONSUMER : L_UBUP_IMemoryConsumer;
	ISVALID : BOOL;
	PTR : POINTER TO BYTE;
	SIZE : UDINT;
END_VAR
END_FUNCTION_BLOCK

METHOD REGISTERCONSUMER
VAR_INPUT
	ITFMEMORYCONSUMER : L_UBUP_IMemoryConsumer;
END_VAR
END_METHOD

METHOD FB_EXIT : BOOL
VAR_INPUT
	BINCOPYCODE : BOOL;
END_VAR
END_METHOD

METHOD FB_INIT : BOOL
VAR_INPUT
	BINITRETAINS : BOOL;
	BINCOPYCODE : BOOL;
END_VAR
END_METHOD

METHOD FB_REINIT : BOOL
END_METHOD

(* ---- L_UBUP_MEMORYPROVIDER1000LREAL.fb ---- *)
FUNCTION_BLOCK L_UBUP_MEMORYPROVIDER1000LREAL EXTENDS L_UBUP_MemoryProvider
VAR
	ALRBUFFER : ARRAY [0..999] OF LREAL;
	PTR : POINTER TO BYTE;
	SIZE : UDINT;
END_VAR
END_FUNCTION_BLOCK

(* ---- L_UBUP_MEMORYPROVIDER100LINT.fb ---- *)
FUNCTION_BLOCK L_UBUP_MEMORYPROVIDER100LINT EXTENDS L_UBUP_MemoryProvider
VAR
	ALINTBUFFER : ARRAY [1..100] OF LINT;
	PTR : POINTER TO BYTE;
	SIZE : UDINT;
END_VAR
END_FUNCTION_BLOCK

(* ---- L_UBUP_MEMORYPROVIDER20LREAL.fb ---- *)
FUNCTION_BLOCK L_UBUP_MEMORYPROVIDER20LREAL EXTENDS L_UBUP_MemoryProvider
VAR
	ALRBUFFER : ARRAY [0..19] OF LREAL;
	PTR : POINTER TO BYTE;
	SIZE : UDINT;
END_VAR
END_FUNCTION_BLOCK

(* ---- L_UBUP_MONITORSTATESERVER.fb ---- *)
FUNCTION_BLOCK L_UBUP_MONITORSTATESERVER
VAR_OUTPUT
	ASCREQUESTPREV : ARRAY [0..c_iMax] OF L_UBUP_MonitorRequest;
	ASCREQUESTPOST : ARRAY [0..c_iMax] OF L_UBUP_MonitorRequest;
	SCREQUESTANNOUNCEDPREV : L_UBUP_MonitorRequest;
	SCREQUESTANNOUNCEDPOST : L_UBUP_MonitorRequest;
	SCREQUESTALTERNATIVEANNOUNCEDPREV : L_UBUP_MonitorRequest;
	SCREQUESTALTERNATIVEANNOUNCEDPOST : L_UBUP_MonitorRequest;
	SCREQUESTACTIVEPREV : L_UBUP_MonitorRequest;
	SCREQUESTACTIVEPOST : L_UBUP_MonitorRequest;
	ISTATE : INT;
END_VAR
VAR
	C_IMAX : INT := 20;
	_ECASE : L_UBUP_StateHandleCase := L_UBUP_StateHandleCase.STATE_POST;
	_IDX1 : INT;
	_IDX2 : INT;
END_VAR
END_FUNCTION_BLOCK

METHOD MONITORCASE
VAR_INPUT
	ECASE : L_UBUP_StateHandleCase;
END_VAR
END_METHOD

METHOD MONITORREQUEST : INT
VAR_INPUT
	ITFREQUEST : L_UBUP_IRequest;
END_VAR
END_METHOD

METHOD MONITORREQUESTANNOUNCED : INT
VAR_INPUT
	ITFREQUESTANNOUNCED : L_UBUP_IRequest;
	ITFREQUESTALTERNATIVE : L_UBUP_IRequest := 0;
	ITFREQUESTACTIVE : L_UBUP_IRequest;
END_VAR
END_METHOD

METHOD REQUESTTOSTRUCT : L_UBUP_MonitorRequest
VAR_INPUT
	ITFREQUEST : L_UBUP_IRequest;
END_VAR
END_METHOD

METHOD RESET : BOOL
END_METHOD

(* ---- L_UBUP_OBJECT.fb ---- *)
FUNCTION_BLOCK L_UBUP_OBJECT
VAR
	_ITFNEXT : L_UBUP_IObject;
	_ITFPREV : L_UBUP_IObject;
	NEXT : L_UBUP_IObject;
	PREV : L_UBUP_IObject;
END_VAR
END_FUNCTION_BLOCK

METHOD CALL_INIT : BOOL
END_METHOD

METHOD SETNEXT : BOOL
VAR_INPUT
	ITFOBJECT : L_UBUP_IObject;
END_VAR
END_METHOD

METHOD SETPREV : BOOL
VAR_INPUT
	ITFOBJECT : L_UBUP_IObject;
END_VAR
END_METHOD

METHOD REQUESTINTERFACE : BOOL
VAR_INPUT
	ID : DINT;
	PITFUNKNOWN : POINTER TO L_UBUP_IUnknown;
END_VAR
END_METHOD

(* ---- L_UBUP_OBJECTQUEUE.fb ---- *)
FUNCTION_BLOCK L_UBUP_OBJECTQUEUE
VAR
	FBSTART : L_UBUP_Object;
	FBFEND : L_UBUP_Object;
	ITFSTART : L_UBUP_IObject := fbStart;
	ITFEND : L_UBUP_IObject := fbfEnd;
	COUNT : DWORD;
	END : L_UBUP_IObject;
	ISEMPTY : BOOL;
	START : L_UBUP_IObject;
END_VAR
END_FUNCTION_BLOCK

METHOD DEQUEUE : BOOL
END_METHOD

METHOD ENQUEUE : BOOL
VAR_INPUT
	ITFOBJECT : L_UBUP_IObject;
END_VAR
END_METHOD

METHOD REMOVE : BOOL
VAR_INPUT
	ITFOBJECT : L_UBUP_IObject;
END_VAR
END_METHOD

METHOD REQUESTINTERFACE : BOOL
VAR_INPUT
	ID : DINT;
	PITFUNKNOWN : POINTER TO L_UBUP_IUnknown;
END_VAR
END_METHOD

METHOD FB_INIT : BOOL
VAR_INPUT
	BINITRETAINS : BOOL;
	BINCOPYCODE : BOOL;
END_VAR
END_METHOD

(* ---- L_UBUP_ONLINECHANGEDETECTION.fb ---- *)
FUNCTION_BLOCK L_UBUP_ONLINECHANGEDETECTION
VAR_OUTPUT
	XONLINECHANGEACTIVE : BOOL;
	DWONLINECHANGECOUNTERPREPARE : DWORD;
	DWONLINECHANGECOUNTERDONE : DWORD;
END_VAR
VAR
	ITFCALLBACK : CmpEventMgr.ICmpEventCallback;
	HINTERFACEPREPAREONLINECHANGE : RTS_IEC_HANDLE;
	HEVENTPREPAREONLINECHANGE : RTS_IEC_HANDLE;
	HINTERFACEONLINECHANGEDONE : RTS_IEC_HANDLE;
	HEVENTONLINECHANGEDONE : RTS_IEC_HANDLE;
END_VAR
END_FUNCTION_BLOCK

METHOD FB_REINIT : BOOL
END_METHOD

METHOD FB_EXIT : BOOL
VAR_INPUT
	BINCOPYCODE : BOOL;
END_VAR
END_METHOD

METHOD FB_INIT : BOOL
VAR_INPUT
	BINITRETAINS : BOOL;
	BINCOPYCODE : BOOL;
END_VAR
END_METHOD

METHOD EVENTCALLBACK : UDINT
VAR_INPUT
	PEVENTPARAM : POINTER TO EventParam;
END_VAR
END_METHOD

METHOD REGISTEREVENT
VAR_INPUT
	XONLYCALLBACKFUNCTION : BOOL;
END_VAR
END_METHOD

METHOD UNREGISTEREVENT
VAR_INPUT
	XONLYCALLBACKFUNCTION : BOOL;
END_VAR
END_METHOD

(* ---- L_UBUP_POOLINSTANCE.fb ---- *)
FUNCTION_BLOCK L_UBUP_POOLINSTANCE EXTENDS L_UBUP_Instance
VAR
	_ITFOWNER : L_UBUP_IFBPool;
	_XWHANDLE : __XWORD;
	_XOCCUPIED : BOOL;
	INSTANCEPTR : POINTER TO BYTE;
	OCCUPIED : BOOL;
END_VAR
END_FUNCTION_BLOCK

METHOD FREE : BOOL
END_METHOD

METHOD OCCUPY : BOOL
VAR_INPUT
	ITFOWNER : L_UBUP_IFBPool;
	XWHANDLE : __XWORD;
END_VAR
END_METHOD

METHOD REQUESTINTERFACE : BOOL
VAR_INPUT
	ID : DINT;
	PITFUNKNOWN : POINTER TO L_UBUP_IUnknown;
END_VAR
END_METHOD

(* ---- L_UBUP_QUEUE.fb ---- *)
FUNCTION_BLOCK L_UBUP_QUEUE
VAR
	_DWPEEKELM : DWORD;
	_DWEMPTYELM : DWORD;
	_DWCOUNTELM : DWORD;
	_DWCAPACITY : DWORD;
	_DWELMSIZE : DWORD;
	COUNT : DWORD;
	ELMSIZE : DWORD;
	ISEMPTY : BOOL;
	ISFULL : BOOL;
END_VAR
END_FUNCTION_BLOCK

METHOD DEQUEUE : BOOL
END_METHOD

METHOD ENQUEUE : BOOL
END_METHOD

METHOD GETEMPTY : BOOL
VAR_OUTPUT
	PBYTE : POINTER TO BYTE;
	DWSIZE : DWORD;
END_VAR
END_METHOD

METHOD GETPEEK : BOOL
VAR_OUTPUT
	PBYTE : POINTER TO BYTE;
	DWSIZE : DWORD;
END_VAR
END_METHOD

METHOD RESET : BOOL
END_METHOD

METHOD FB_INIT : BOOL
VAR_INPUT
	BINITRETAINS : BOOL;
	BINCOPYCODE : BOOL;
END_VAR
END_METHOD

METHOD GETELMPTR : POINTER TO BYTE
VAR_INPUT
	DWELMIDX : DWORD;
END_VAR
END_METHOD

METHOD GETQUEUEINFO
VAR_OUTPUT
	DWCAPACITY : DWORD;
	DWELMSIZE : DWORD;
END_VAR
END_METHOD

(* ---- L_UBUP_QUEUEARRAYCONTROL.fb ---- *)
FUNCTION_BLOCK L_UBUP_QUEUEARRAYCONTROL
VAR_OUTPUT
	DWCAPACITY : DWORD;
	DWCOUNTELM : DWORD;
	DWFIRSTELM : DWORD;
	DWLASTELM : DWORD;
	DWACTIVEELM : DWORD;
END_VAR
VAR
	COUNT : DWORD;
	ELMSIZE : DWORD;
	ISEMPTY : BOOL;
	ISFULL : BOOL;
END_VAR
END_FUNCTION_BLOCK

METHOD DEQUEUE : BOOL
END_METHOD

METHOD DEQUEUELAST : BOOL
END_METHOD

METHOD ENQUEUE : BOOL
END_METHOD

METHOD GETEMPTY : BOOL
VAR_OUTPUT
	PBYTE : POINTER TO BYTE;
	DWSIZE : DWORD;
END_VAR
END_METHOD

METHOD GETPEEK : BOOL
VAR_OUTPUT
	PBYTE : POINTER TO BYTE;
	DWSIZE : DWORD;
END_VAR
END_METHOD

METHOD RESET : BOOL
END_METHOD

METHOD FB_INIT : BOOL
VAR_INPUT
	BINITRETAINS : BOOL;
	BINCOPYCODE : BOOL;
	DWCAPACITY : DWORD;
END_VAR
END_METHOD

METHOD LOADCAPACITY : BOOL
VAR_INPUT
	DWCAPACITY : DWORD;
END_VAR
END_METHOD

(* ---- L_UBUP_REQUESTTRANSITION.fb ---- *)
FUNCTION_BLOCK L_UBUP_REQUESTTRANSITION
VAR_INPUT
	XENABLE : BOOL := TRUE;
	XREQUEST : BOOL;
END_VAR
VAR_OUTPUT
	XREQUESTACTIVE : BOOL;
	IACTUALPRIO : INT := L_UBUP_Internal.g_iLowestRequestPrio;
	XCONDITIONVERIFY : BOOL;
END_VAR
VAR
	_ITFCONDITION : L_UBUP_ICondition;
	_ITFSTATESERVER : L_UBUP_IStateServer;
	_ITFSTATECLIENT : L_UBUP_IStateClient;
	_ITFREQUEST_THIS : L_UBUP_IRequest := THIS^;
	_ETARGETSTATE : INT;
	_IPRIO : INT;
	_XEDGEREQUESTFORCEENTRY : BOOL;
	_XEDGEUP : BOOL;
	_XEDGEDOWN : BOOL;
	_XREQUEST_OLD : BOOL;
	_XENABLE_OLD : BOOL;
	ACTUALPRIO : INT;
	ACTUALSTATE : INT;
	CONDITIONVALID : BOOL;
	REQUESTACTIVE : BOOL;
	REQUESTEDGEDOWN : BOOL;
	REQUESTEDGEUP : BOOL;
	REQUESTLEVEL : BOOL;
END_VAR
END_FUNCTION_BLOCK

METHOD VERIFY : BOOL
VAR_OUTPUT
	XCONDITIONERROR : BOOL;
	EERRORIDPROPOSED : L_IE1P_Error;
END_VAR
END_METHOD

METHOD CONFIRM : INT
VAR_IN_OUT
	IREQUEST : L_UBUP_IRequest;
END_VAR
END_METHOD

METHOD FORCESTATEENTRY : BOOL
END_METHOD

METHOD FB_INIT : BOOL
VAR_INPUT
	BINITRETAINS : BOOL;
	BINCOPYCODE : BOOL;
	ITFSTATESERVER : L_UBUP_IStateServer;
	ITFCONDITION : L_UBUP_ICondition;
	IPRIO : INT;
	ETARGETSTATE : INT;
	XEDGEREQUESTFORCEENTRY : BOOL;
END_VAR
END_METHOD

METHOD EDGEUPIMPL : BOOL
END_METHOD

METHOD RESET
END_METHOD

(* ---- L_UBUP_REQUESTTRANSITIONEDGE.fb ---- *)
FUNCTION_BLOCK L_UBUP_REQUESTTRANSITIONEDGE EXTENDS L_UBUP_RequestTransition
VAR
	XCONDITIONERROR : BOOL;
	ECONDITIONERRORID : L_IE1P_Error;
END_VAR
END_FUNCTION_BLOCK

METHOD FORCESTATEENTRY : BOOL
END_METHOD

(* ---- L_UBUP_REQUESTTRANSITIONLEVEL.fb ---- *)
FUNCTION_BLOCK L_UBUP_REQUESTTRANSITIONLEVEL EXTENDS L_UBUP_RequestTransition
VAR
	_XVERIFYRTRIG : BOOL;
END_VAR
END_FUNCTION_BLOCK

METHOD FORCESTATEENTRY : BOOL
END_METHOD

METHOD VERIFY : BOOL
VAR_OUTPUT
	XCONDITIONERROR : BOOL;
	EERRORIDPROPOSED : L_IE1P_Error;
END_VAR
END_METHOD

(* ---- L_UBUP_STATECLIENTPROXY.fb ---- *)
FUNCTION_BLOCK L_UBUP_STATECLIENTPROXY
VAR_INPUT
	ITFDECORATOR : L_UBUP_IStateClientDecorator;
END_VAR
VAR
	_ITFCLIENT : L_UBUP_IStateClient;
	_ITFALLOCPOINTADRPROVIDER : L_UBUP_IAllocPointAdrProvider;
END_VAR
END_FUNCTION_BLOCK

METHOD ALLOCPOINTADR
VAR_OUTPUT
	IERRORID : INT;
END_VAR
END_METHOD

METHOD CALLFBS
VAR_INPUT
	ECASE : L_UBUP_StateHandleCase;
END_VAR
END_METHOD

METHOD CALLSTATE
VAR_INPUT
	ITFSTATESERVER : L_UBUP_IStateServer;
	ISTATE : INT;
	ECASE : L_UBUP_StateHandleCase;
END_VAR
END_METHOD

METHOD CHECKTRANSITION
VAR_INPUT
	ITFSTATESERVER : L_UBUP_IStateServer;
END_VAR
END_METHOD

METHOD DISABLECLIENT : BOOL
VAR_INPUT
	XFIRSTCALL : BOOL;
END_VAR
END_METHOD

METHOD ENABLECLIENT : BOOL
VAR_INPUT
	XFIRSTCALL : BOOL;
END_VAR
END_METHOD

METHOD FINALIZECYCLE
END_METHOD

METHOD LEAVESTATE
END_METHOD

METHOD PREPARECYCLE
END_METHOD

METHOD PREPARESTATECHANGE
END_METHOD

METHOD STIMULATETRANSITION
VAR_INPUT
	ECASE : L_UBUP_StateHandleCase;
END_VAR
END_METHOD

METHOD UPDATECONDITIONERROR : BOOL
VAR_INPUT
	ITFREQUEST : L_UBUP_IRequest;
END_VAR
END_METHOD

METHOD REQUESTINTERFACE : BOOL
VAR_INPUT
	ID : DINT;
	PITFUNKNOWN : POINTER TO L_UBUP_IUnknown;
END_VAR
END_METHOD

METHOD FB_INIT : BOOL
VAR_INPUT
	BINITRETAINS : BOOL;
	BINCOPYCODE : BOOL;
	ITFCLIENT : L_UBUP_IStateClient;
END_VAR
END_METHOD

(* ---- L_UBUP_STATESERVER.fb ---- *)
FUNCTION_BLOCK L_UBUP_STATESERVER
VAR_INPUT
	XENABLE : BOOL;
END_VAR
VAR_OUTPUT
	XBUSY : BOOL;
	XACTIVE : BOOL;
	XERROR : BOOL;
	EERRORID : L_IE1P_Error;
	ESTATEACTUAL : INT := -1;
END_VAR
VAR
	_ITFREQUESTACTIVE : L_UBUP_IRequest;
	_ITFREQUESTANNOUNCED : L_UBUP_IRequest;
	_ITFCLIENT : L_UBUP_IStateClient;
	_ITFALLOCPOINTADRPROVIDER : L_UBUP_IAllocPointAdrProvider;
	_ITFALTERNATIVEREQUESTBYFAILEDCONDITION : L_UBUP_IAlternativeRequestByFailedCondition;
	_ITFMONITOR : L_UBUP_IMonitorStateServer;
	_ESTATEPREV : INT := -1;
	_XCONDITIONERRORTMP : BOOL;
	_ECONDITIONERRORIDTMP : L_IE1P_Error;
	_XENABLEOLD : BOOL;
	_XFREEZEREQUEST : BOOL;
	_IFREEZEREQUESTPRIO : INT := 10;
	_EERRORIDBYBLOCKEFREEZEREQUEST : L_IE1P_Error;
	_XANNOUNCENEWREQUEST : BOOL;
	_IERRORID : INT;
	ACTUALCLIENT : L_UBUP_IStateClient;
	ACTUALSTATE : INT;
	FREEZEREQUESTACTIVE : BOOL;
	IFREEZEREQUESTPRIO : INT;
	ITFALTERNATIVEREQUESTBYFAILEDCONDITION : L_UBUP_IAlternativeRequestByFailedCondition;
	MONITORSTATESERVER : L_UBUP_IMonitorStateServer;
END_VAR
END_FUNCTION_BLOCK

METHOD ANNOUNCENEWREQUEST
END_METHOD

METHOD FREEZEREQUEST
VAR_INPUT
	EERRORIDBYBLOCKEFREEZEREQUEST : L_IE1P_Error;
END_VAR
END_METHOD

METHOD ISACTIVE : BOOL
VAR_INPUT
	ITFREQUEST : L_UBUP_IRequest;
END_VAR
END_METHOD

METHOD REQUESTS : INT
VAR_INPUT
	ITFREQUEST : L_UBUP_IRequest;
END_VAR
END_METHOD

METHOD UNFREEZEREQUEST : BOOL
END_METHOD

METHOD VERIFYFREEZEREQUEST : BOOL
VAR_INPUT
	ITFREQUEST : L_UBUP_IRequest;
END_VAR
VAR_OUTPUT
	XCONDITIONERROR : BOOL;
	EERRORIDPROPOSED : L_IE1P_Error;
END_VAR
END_METHOD

METHOD FB_INIT : BOOL
VAR_INPUT
	BINITRETAINS : BOOL;
	BINCOPYCODE : BOOL;
	ITFCLIENT : L_UBUP_IStateClient;
END_VAR
END_METHOD

METHOD EXECUTEREQUESTANNOUNCED
END_METHOD

(* ---- L_UBUP_STRINGCOLLECTIONWRITER.fb ---- *)
FUNCTION_BLOCK L_UBUP_STRINGCOLLECTIONWRITER EXTENDS L_UBUP_FreeRunTask
VAR_INPUT
	ITFSTRINGS : L_UBUP_IStringCollection;
	STRFILENAME : STRING(255);
	STRFILEPATH : STRING(255);
END_VAR
END_FUNCTION_BLOCK

METHOD STARTACTION
VAR_OUTPUT
	XCOMPLETE : BOOL;
	IERRORID : INT;
END_VAR
END_METHOD

METHOD FB_INIT : BOOL
VAR_INPUT
	BINITRETAINS : BOOL;
	BINCOPYCODE : BOOL;
END_VAR
END_METHOD

METHOD EXECUTEIMPL : UDINT
END_METHOD

(* ---- L_UBUP_STRINGQUEUE.fb ---- *)
FUNCTION_BLOCK L_UBUP_STRINGQUEUE EXTENDS L_UBUP_Queue
VAR
	ASTRLINES : ARRAY [1..c_LineCount] OF STRING(255);
	C_LINECOUNT : DWORD := 100;
END_VAR
END_FUNCTION_BLOCK

METHOD GETELMPTR : POINTER TO BYTE
VAR_INPUT
	DWELMIDX : DWORD;
END_VAR
END_METHOD

METHOD GETQUEUEINFO
VAR_OUTPUT
	DWCAPACITY : DWORD;
	DWELMSIZE : DWORD;
END_VAR
END_METHOD

(* ---- L_UBUP_SYMBOLCONFIG.fb ---- *)
FUNCTION_BLOCK L_UBUP_SYMBOLCONFIG
VAR
	_VARACCESSIBASE : IecVarAccessLibrary.IBase;
	_PPIVARACCESS3 : POINTER TO IecVarAccessLibrary.IIecVarAccess3;
	_VARACCESS3 : IecVarAccessLibrary.IIecVarAccess3;
	_PPIVARACCESS4 : POINTER TO IecVarAccessLibrary.IIecVarAccess4;
	_VARACCESS4 : IecVarAccessLibrary.IIecVarAccess4;
	_PPIVARACCESS5 : POINTER TO IecVarAccessLibrary.IIecVarAccess5;
	_VARACCESS5 : IecVarAccessLibrary.IIecVarAccess5;
	_SSYMBOL : STRING(255);
	_HNODE : IecVarAccessLibrary.ICollections.IBaseTreeNode;
	_VARINFO : VariableInformationStruct;
END_VAR
END_FUNCTION_BLOCK

METHOD FINDSYMBOL : RTS_IEC_RESULT
VAR_INPUT
	HNODE : IecVarAccessLibrary.ICollections.IBaseTreeNode;
	XWADDRESS : __XWORD;
END_VAR
VAR_IN_OUT
	SSYMBOL : STRING(255);
END_VAR
END_METHOD

METHOD GETADDRESS : POINTER TO BYTE
VAR_OUTPUT
	RESULT : RTS_IEC_RESULT;
END_VAR
END_METHOD

METHOD GETSIZE : __XWORD
VAR_OUTPUT
	RESULT : RTS_IEC_RESULT;
END_VAR
END_METHOD

METHOD GETSYMBOL : STRING
VAR_OUTPUT
	RESULT : RTS_IEC_RESULT;
END_VAR
END_METHOD

METHOD GETVARSTRING : BOOL
VAR_OUTPUT
	SVALUE : STRING;
END_VAR
END_METHOD

METHOD GETVARTYPE : BOOL
VAR_OUTPUT
	EVARTYPE : L_UBUP_VarType;
END_VAR
END_METHOD

METHOD GETVARVALUE : BOOL
VAR_OUTPUT
	EVARTYPE : L_UBUP_VarType;
	UVARVALUE : L_UBUP_VarValue;
END_VAR
END_METHOD

METHOD GETVARVALUEASDWORD : BOOL
VAR_OUTPUT
	DWVALUE : DWORD;
END_VAR
END_METHOD

METHOD GETVARVALUEASLINT : BOOL
VAR_OUTPUT
	LIVALUE : LINT;
END_VAR
END_METHOD

METHOD GETVARVALUEASLREAL : BOOL
VAR_OUTPUT
	LRVALUE : LREAL;
END_VAR
END_METHOD

METHOD GETVARVALUEASWORD : BOOL
VAR_OUTPUT
	WVALUE : WORD;
END_VAR
END_METHOD

METHOD GETVARIABLE : BOOL
VAR_OUTPUT
	SCVARIABLE : L_UBUP_Variable;
END_VAR
END_METHOD

METHOD INIT : BOOL
VAR_IN_OUT
	RESULT : RTS_IEC_RESULT;
END_VAR
END_METHOD

METHOD REQUEST : BOOL
VAR_INPUT
	SSYMBOL : STRING(255);
END_VAR
END_METHOD

(* ---- L_UBUP_TIMINGCONTROLLER.fb ---- *)
FUNCTION_BLOCK L_UBUP_TIMINGCONTROLLER
VAR
	_STARTOPTIME_US : SYSTIME;
	_STARTINVTIME_US : SYSTIME;
	_CURRENTTIME_US : SYSTIME;
	_TIMELIMIT_US : SYSTIME;
	_TIMEOUT_US : SYSTIME;
	TIMELIMIT : SYSTIME;
	TIMEOUT : SYSTIME;
END_VAR
END_FUNCTION_BLOCK

METHOD CHECKTIMING
VAR_OUTPUT
	XTIMEOUT : BOOL;
	XTIMELIMIT : BOOL;
END_VAR
END_METHOD

METHOD STARTINVOCATIONTIMER
END_METHOD

METHOD STARTOPERATIONTIMER
END_METHOD

(* ---- L_UBUP_TRACEARRAY.fb ---- *)
FUNCTION_BLOCK L_UBUP_TRACEARRAY
VAR_INPUT
	ALRDATA : POINTER TO LREAL;
	XEXECUTE : BOOL;
	XABORT : BOOL;
END_VAR
VAR_OUTPUT
	XDONE : BOOL;
	XBUSY : BOOL;
	XACTIVE : BOOL;
	XCOMMANDABORTED : BOOL;
	XERROR : BOOL;
	EERRORID : L_IE1P_Error;
	LRACTUALVALUE : LREAL;
END_VAR
VAR
	_DWMININDEX : DWORD;
	_DWMAXINDEX : DWORD;
	_DWACTINDEX : DWORD;
	_MODEL : L_UBUP_BehaviourModel_ETrigA;
END_VAR
END_FUNCTION_BLOCK

METHOD CYCLICACTION
VAR_INPUT
	ITFTIMINGCONTROLLER : L_UBUP_ITimingController;
END_VAR
VAR_OUTPUT
	XCOMPLETE : BOOL;
	XABORT : BOOL;
	IERRORID : INT;
END_VAR
END_METHOD

METHOD FINALIZEACTION
VAR_INPUT
	XABORTPROPOSED : BOOL;
	IERRORIDPROPOSED : INT;
END_VAR
VAR_OUTPUT
	XCOMPLETE : BOOL;
	XABORT : BOOL;
	IERRORID : INT;
END_VAR
END_METHOD

METHOD RESETACTION
VAR_OUTPUT
	XCOMPLETE : BOOL;
END_VAR
END_METHOD

METHOD STARTACTION
VAR_OUTPUT
	XCOMPLETE : BOOL;
	IERRORID : INT;
END_VAR
END_METHOD

(* ---- L_UBUP_VENDORIDCHECKER.fb ---- *)
FUNCTION_BLOCK L_UBUP_VENDORIDCHECKER
VAR_OUTPUT
	DWVENDORID : DWORD;
END_VAR
END_FUNCTION_BLOCK

METHOD PERFORMCHECK : BOOL
VAR_INPUT
	WCONTEXT : DWORD;
END_VAR
END_METHOD

METHOD REQUESTINTERFACE : BOOL
VAR_INPUT
	ID : DINT;
	PITFUNKNOWN : POINTER TO L_UBUP_IUnknown;
END_VAR
END_METHOD
